IF bReset
     AND bError
THEN
	udnErrorNo := 0;					(* Error number *)
	sErrorMsg := ''; 					(* Error message *)
	tonWatchDog(IN := FALSE);

END_IF

(* Check inputs  *)
rtHandOn(CLK := bHandOn);
rtAutoOn(CLK := bAutoOn AND bReleaseOn AND bReleasePowerOn);
rtAutoOff(CLK := bAutoOff);

(* Check operating mode *)
IF bAutoHand					(* Automatic *)
THEN
	IF rtAutoOff.Q
	THEN
		bPowerOn := FALSE;

	ELSIF rtAutoOn.Q
		    AND bReleasePowerOn
	THEN
		bPowerOn := TRUE;
	END_IF;

ELSE						(* Manual *)
	IF rtHandOn.Q
	THEN
		IF bPowerOn
		THEN
			bPowerOn := FALSE;

		ELSIF bReleaseOn
			   AND bReleasePowerOn
		THEN
			bPowerOn := TRUE;
		END_IF
	END_IF

END_IF;

(* Timer starts when cylinder is not  in base and work position *)
tonWatchDog(
	IN := bPowerOn
		 AND bPowerSupplyOn
		 AND NOT bReady,
	PT := tTimeOut + tReadyDelay
);

(* Error if cylinder does not reach base or work position*)
IF tonWatchDog.Q
   AND NOT bError
THEN
	IF bPowerOn AND NOT bReady
	THEN
		udnErrorNo := 1; 								(* Set error number *)
		sErrorMsg := 'Not ready error';
	END_IF
END_IF

tonPowerSupplyOn(
	IN := bNoEStop
		 AND NOT bPowerSupplyOn,
	PT := tTimeOut
);

IF tonPowerSupplyOn.Q
THEN
	udnErrorNo := 2; 								(* Set error number *)
	sErrorMsg := 'Power supply error';
END_IF
(*
IF lrSetTemp > 0
     AND lrActTemp > lrMaxTemp
THEN
	udnErrorNo := 2; 								(* Set error number *)
	sErrorMsg := 'Temperatur over range';
END_IF
*)

bError := udnErrorNo <> 0;

fbReadyDelay(
	bEnable := TRUE,
	bIn := bPowerOn,
	tDelay := tReadyDelay
);

IF lrSetTemp <> 0
     AND bAutoHand 			(* Automatic *)
THEN
	bReady := bPowerOn
			   AND lrActTemp >= lrSetTemp;
ELSE
	bReady := fbReadyDelay.bOut;
END_IF

(* Scaling power *)
fbScalingSP(
	bEnable := TRUE,
	lrInput := lrSPPower, (* [%] *)
	lrXLowLimit := 0, (* [%] *)
	lrXUpperLimit := 100, (* [%] *)
	lrYLowLimit := lrPowerMin, (* 16#0000 = 0 [V] *)
	lrYUpperLimit := lrPowerMax, (* 16#7FFF = 10 [V] *)
	usiPrecision := 2
);
unCVPower := LREAL_TO_UINT(fbScalingSP.lrOutputPV);

END_FUNCTION_BLOCK

// ---- POUs/Tc2 Objects/Automation/NCiChannel/FB_CfgAxisInExt3DGroup.TcPOU
FUNCTION_BLOCK FB_CfgAxisInExt3DGroup
(*

The function block used to detects if are axis in a group or if the group is occupied. 

Constructor: 		Patryk Panylo
Company:		E. Riexinger GmbH
Date:			23.04.2015
Version:			1.00

Date:			Revision:		Who:				Comment
dd.mm.yyyy		x.xx			Initials			comment

*)
VAR_INPUT
	(* Input variables / Eingang Variablen *)
	bEnable						:BOOL;			(* Signal FB enable *)
	bExecute					:BOOL; 			(* Execute the programm *)
	udnGrpId						:UDINT;			(* Id of the 3D Group *)
	tTimeOut						:TIME := T#5s;	(* TimeOut *)
END_VAR
VAR_OUTPUT
	(* Output variables / Ausgang Variablen *)
	bGrpOccupied				:BOOL;			(* Axis in group detected *)
	bGrpEmpty					:BOOL;			(* Axis not in group detected *)
	bDone						:BOOL;			(* Command done *)
	bBusy						:BOOL;			(* Command busy *)
	bError						:BOOL;			(* Command error  *)
	udnErrorNo					:UDINT;			(* Error number *)
	sErrorMsg					:STRING; 		(* Error message *)
END_VAR
VAR_IN_OUT
	(* Input Output variables / Ausgang Variablen *)

END_VAR
VAR
	(* Enummerations *)
	etCfgAxisInExt3DGrp			:ET_CfgAxisInExt3DGroup;

	(* Variables *)
	stExt3dGrp 					:NCI_EXT3DGROUP;				(* Contains the Axis ID's *)

	bFirstTime					:BOOL;

	(* References *)

	(* Interfaces *)

	(* Instances *)
	fbCfgReadExt3DAxisIds		:CfgReadExt3DAxisIds;				(* The block CfgReadExt3DAxisIds reads the axis configuration of the advanced 3D group. *)

END_VAR

IF NOT bEnable
THEN
	bGrpOccupied := FALSE;			(* Axis in group detected *)
	bGrpEmpty :=FALSE;				(* Axis not in group detected *)
	bDone := FALSE;					(* Program done *)
	bBusy := FALSE;                                  	(* Program not busy *)
	bError := FALSE;                                 	(* Program not error *)
	udnErrorNo := 0;					(* Error number *)
	sErrorMsg := ''; 					(* Error message *)

	bFirstTime := FALSE;
	RETURN;
END_IF;

IF NOT bFirstTime
THEN
	bGrpOccupied := FALSE;			(* Axis in group detected *)
	bGrpEmpty :=FALSE;				(* Axis not in group detected *)
	bDone := FALSE;                                 	(* Program done *)
	bBusy := FALSE;                                  	(* Program not busy *)
	bError := FALSE;                                 	(* Program not error *)
	udnErrorNo := 0;					(* Error number *)
	sErrorMsg := ''; 					(* Error message *)

	fbCfgReadExt3DAxisIds(
		bExecute := FALSE,
		stExt3dGroup := stExt3dGrp
	);

	etCfgAxisInExt3DGrp := ET_CfgAxisInExt3DGrp_eWaitExecute;       				(* Next step *)
	
	bFirstTime := TRUE;
END_IF;

CASE etCfgAxisInExt3DGrp OF
        
	ET_CfgAxisInExt3DGrp_eWaitExecute:
		bBusy := FALSE;                                     		(* Program not busy *)
		bError := FALSE;                                    		(* Program not error *)

		IF bExecute
		THEN
			bDone := FALSE;                                 	(* Program done, in position *)
			bBusy := TRUE;                                  	(* Program busy *)
			udnErrorNo := 0;					(* Error number *)
			sErrorMsg := ''; 					(* Error message *)
	           
			etCfgAxisInExt3DGrp := ET_CfgAxisInExt3DGrp_eReadExt3DAxisIds;         		(* Next step *)
		END_IF;

	ET_CfgAxisInExt3DGrp_eReadExt3DAxisIds:

		fbCfgReadExt3DAxisIds(			(* Read axis ID's *)
			bExecute := TRUE ,
			nGroupId := udnGrpId,
			tTimeOut := tTimeOut,
			stExt3dGroup := stExt3dGrp
		);

		IF NOT fbCfgReadExt3DAxisIds.bBusy
		     AND NOT fbCfgReadExt3DAxisIds.bErr
		THEN
			fbCfgReadExt3DAxisIds(
				bExecute := FALSE,
				stExt3dGroup := stExt3dGrp
			);

			bGrpEmpty :=	stExt3dGrp.nXAxisId = 0						(* Check if axis in Group *)
						AND stExt3dGrp.nYAxisId = 0
						AND stExt3dGrp.nZAxisId = 0
						AND stExt3dGrp.nQ1AxisId =  0
						AND stExt3dGrp.nQ2AxisId =  0
						AND stExt3dGrp.nQ3AxisId =  0
						AND stExt3dGrp.nQ4AxisId =  0
						AND stExt3dGrp.nQ5AxisId =  0;
			bGrpOccupied := NOT bGrpEmpty ;
			
			etCfgAxisInExt3DGrp := ET_CfgAxisInExt3DGrp_eDone;            			(* Next step *)

		ELSIF fbCfgReadExt3DAxisIds.bErr
		THEN
			udnErrorNo := fbCfgReadExt3DAxisIds.nErrId;						(* Set error number *)

			fbCfgReadExt3DAxisIds(
				bExecute := FALSE,
				stExt3dGroup := stExt3dGrp
			);

			etCfgAxisInExt3DGrp := ET_CfgAxisInExt3DGrp_eError;            			(* Next step *)
		
		END_IF

	ET_CfgAxisInExt3DGrp_eDone:
		bDone := TRUE;                                      		(* Program done, in position *)
		bBusy := FALSE;                                     		(* Program not busy *)
	
		etCfgAxisInExt3DGrp := ET_CfgAxisInExt3DGrp_eNoExecute;            		(* Next step *)
	
	ET_CfgAxisInExt3DGrp_eError:
		bDone := FALSE;                                    	 	(* Program done, in position *)
		bError := TRUE;                                     		(* Program error *)
		bBusy := FALSE;                                     		(* Program not busy *)

		etCfgAxisInExt3DGrp := ET_CfgAxisInExt3DGrp_eNoExecute;            		(* Next step *)
	
	ET_CfgAxisInExt3DGrp_eNoExecute:
		IF NOT bExecute
		THEN
			bDone := FALSE;                                 	(* Program done *)
			bBusy := FALSE;                                 	(* Program not busy *)
			bError := FALSE;                                		(* Program not error *)

			etCfgAxisInExt3DGrp := ET_CfgAxisInExt3DGrp_eWaitExecute;       		(* Next step *)
	
		END_IF;
        
END_CASE;

END_FUNCTION_BLOCK

// ---- POUs/Tc2 Objects/Automation/Sawband/FB_Sawband.TcPOU
FUNCTION_BLOCK FB_Sawband
(*

The function block used to control the saw.

Constructor: 		Patryk Panylo
Company:		E. Riexinger GmbH
Date:			04.11.2015
Version:			1.00

Date:			Revision:		Who:				Comment
dd.mm.yyyy		x.xx			Initials			comment

*)
VAR_INPUT
	(* Input variables / Eingang Variablen *)
	bEnable					:BOOL;						(* Enable FB signal *)
	bNoEStop				:BOOL;						(* No ermergency Stop / Keine Notaus *)
	bAirPressure				:BOOL;						(* Signal air pressure *)
	bAutoHand				:BOOL;						(* Auto := TRUE, Hand := FALSE *)
	bHandStart				:BOOL;						(* Sawband hand start *)
	bHandStop				:BOOL;						(* Sawband hand stop *)
	bAutoStart				:BOOL;						(* Sawband auto start *)
	bAutoStop				:BOOL;						(* Sawband auto stop *)
	bSawbandAir				:BOOL;						(* Sawband air on *)
	bSawbandCtrlOK			:BOOL;						(* Sawband controller ok *)
	bSawbandNOK			:BOOL;						(* Sawband error *)
	udnIncEnc				:UDINT;						(* Value of encoder increment *)
	udnScalingDenom			:UDINT := 1;	  				(* Denominator for the conversion factor at the conversion of bus data to technical units [INC] *)
	lrScalingNum				:LREAL := 1.0;  				(* Numerator for the conversion factor at the conversion of bus data to technical units [technical units] *)
	lrTaskCycle				:LREAL := 0.002;				(* Cycle time of the task [sec], 0.002[s] => 2ms *)
	lrSawbandRefVelo		:LREAL := 1.0;					(* Referenc velocity of sawband [technical units/s]*)
	tSawbandCtrlOnDelay		:TIME := t#3s;					(* Sawband on delay *)
	tSawbandAirOffDelay		:TIME := t#10s;				(* Sawband air off delay *)
	tSawbandReadyDelay		:TIME := t#5s;					(* Sawband ready delay *)
END_VAR
VAR_OUTPUT
	(* Output variables / Ausgang Variablen *)
	bSawbandReady			:BOOL;						(* Sawband ready *)
	bSawbandCtrlOn			:BOOL;						(* Sawband controller on *)
	bSawbandAirOn			:BOOL;						(* Sawband air on*)
	bNotMoving				:BOOL;						(* Axis not moving *)
	lrActPosition				:LREAL;						(* Actual position [mm] *)
	lrActVelocity				:LREAL;						(* Actual velocity [mm/s] *)
	bError					:BOOL;						(* Error *)
	udnErrorNo				:UDINT;
	udnMessageNo			:UDINT;
	sMsg					:STRING;
END_VAR
VAR_IN_OUT

END_VAR
VAR
	(* Enummerations *)

	(* Variables *)
	stEncoderConfig				:ST_EncoderConfig;			(* Encoder configuration *)
	stAxis						:ST_AXIS_REF_V2;			(* The AXIS_REF data type  is an interface between the PLC and the NC and contains axis information *)
	bFirstTime					:BOOL;						(* First cycle *)

	(* References *)

	(* Interfaces *)

	(* Instances *)
	rtHandStart				:R_TRIG;
	rtHandStop				:R_TRIG;
	rtAutoStart				:R_TRIG;
	rtAutoStop				:R_TRIG;
	tonSawbandCtrlOnDelay	:TON;						(* Timer to delay *)
	tofSawbandAirOffDelay		:TOF;						(* Timer to delay *)
	tonSawbandReadyDelay  	:TON;						(* Timer to delay *)

	fbPositionEncoder			:FB_PositionEncoder;
END_VAR

IF NOT bEnable
THEN
	bSawbandCtrlOn := FALSE;
	bSawbandAirOn := FALSE;
	bError := FALSE;
	udnErrorNo := 0;
	udnMessageNo := 0;
	sMsg := '';
	tonSawbandCtrlOnDelay(IN := FALSE,
					       	    PT := tSawbandCtrlOnDelay);
	tofSawbandAirOffDelay(IN := FALSE,
	            			 	 PT := tSawbandAirOffDelay);
	tonSawbandReadyDelay(IN := FALSE,
					       		PT := tSawbandReadyDelay);
	bFirstTime := FALSE;
    RETURN;
END_IF;

IF NOT bFirstTime
THEN
	bError := FALSE;
	udnErrorNo := 0;
	udnMessageNo := 0;
	sMsg := '';
	tonSawbandCtrlOnDelay(IN := FALSE,
					       	    PT := tSawbandCtrlOnDelay);
	tofSawbandAirOffDelay(IN := FALSE,
	            			 	 PT := tSawbandAirOffDelay);
	tonSawbandReadyDelay(IN := FALSE,
					       		PT := tSawbandReadyDelay);
	bFirstTime := TRUE;
END_IF;

(* Start / Stop sawband *)
rtHandStart(CLK := bHandStart);
rtHandStop(CLK := bHandStop);
rtAutoStart(CLK := bAutoStart);
rtAutoStop(CLK := bAutoStop);

IF rtHandStop.Q
     OR rtAutoStop.Q
     OR NOT bNoEStop
     OR bSawbandNOK
THEN
	tofSawbandAirOffDelay.IN := FALSE;;
	tonSawbandCtrlOnDelay.IN := FALSE;

ELSIF SEL(bAutoHand, rtHandStart.Q, rtAutoStart.Q)
	    AND bNoEStop
	    AND bAirPressure
	    AND NOT bSawbandNOK
THEN
	tofSawbandAirOffDelay.IN := TRUE;;
	tonSawbandCtrlOnDelay.IN := TRUE;

END_IF

(* Sawband air stop after delay *)
tofSawbandAirOffDelay(
         PT := tSawbandAirOffDelay
);

bSawbandAirOn := tofSawbandAirOffDelay.Q
				OR ( NOT bAutoHand
					AND bSawbandAir);

(* Sawband controller on after delay *)
tonSawbandCtrlOnDelay(
         PT := tSawbandCtrlOnDelay
);

bSawbandCtrlOn := tonSawbandCtrlOnDelay.Q;

(* Sawband ready after delay *)
tonSawbandReadyDelay(
	IN := bSawbandCtrlOn,
	PT := tSawbandReadyDelay
);

A_PositionDynamics();
A_Alarm();

bSawbandReady := bSawbandCtrlOK
				   AND NOT bSawbandNOK
				   AND NOT bNotMoving
				   AND NOT bError
				   AND lrActVelocity >= lrSawbandRefVelo
				   AND tonSawbandReadyDelay.Q;

ACTION A_Alarm:

(* Check error *)
IF bSawbandNOK
THEN
	udnErrorNo := 1;
	udnMessageNo := 0;
	sMsg := 'Sawband nok signal';

ELSIF (NOT bSawbandCtrlOK
	    	      OR bNotMoving)
	   AND tonSawbandReadyDelay.Q
THEN
	udnErrorNo := 2;
	udnMessageNo := 0;
	sMsg := 'Sawband not ready';

ELSE
	udnErrorNo := 0;
	udnMessageNo := 0;
	sMsg := '';

END_IF

bError := udnErrorNo > 0;
END_ACTION

ACTION A_PositionDynamics:

(* Position encoding *)
stEncoderConfig.etScalingMethod := ET_ScalingMethod_eSMLinear;
stAxis.stScaling.etScalingMethod := ET_ScalingMethod_eSMLinear;
stAxis.stScaling.lrTaskCycle := lrTaskCycle;
stAxis.stScaling.udnScalingDenom := udnScalingDenom; (* inc *)
stAxis.stScaling.lrScalingNum := lrScalingNum; (* mm *)

fbPositionEncoder(
	bEnable := TRUE,
	dwEncCurrentValue := udnIncEnc,
	stEncCfg := stEncoderConfig,
	pAxis := ADR(stAxis)
);

lrActPosition := fbPositionEncoder.pAxis^.stPosition.lrActPos / 1000 (* m *);
lrActVelocity := fbPositionEncoder.pAxis^.stDynamics.lrActVelo * 60 (* mm/min *);

bNotMoving := FALSE;

IF lrActVelocity = 0.0
THEN
	bNotMoving := TRUE;
END_IF
END_ACTION

END_FUNCTION_BLOCK

// ---- POUs/Tc2 Objects/Automation/Spindle/FB_CoolingDevice.TcPOU
FUNCTION_BLOCK FB_CoolingDevice
(*

The function block used to control power supply.

Constructor: 		Patryk Panylo
Company:		E. Riexinger GmbH
Date:			23.04.2015
Version:			1.00

Date:			Revision:		Who:				Comment
dd.mm.yyyy		x.xx			Initials			comment

*)
VAR_INPUT
	(* Input variables / Eingang Variablen *)
	bEnable					:BOOL;						(* Enable FB signal *)
	bIn						:BOOL;						(* Input signal *)
	tCoolingDeviceOn			:TIME := t#2s;					(* Timeout power supply on *)
	tCoolingDeviceOff			:TIME := t#1s;					(* Timeout power supply off *)
END_VAR
VAR_OUTPUT
	(* Output variables / Ausgang Variablen *)
	bOut					:BOOL;						(* Air pressure ok *)
	bError					:BOOL;						(* Error by no air pressure *)
	udnErrorNo				:UDINT;
	udnMessageNo			:UDINT;
	sMsg					:STRING;
END_VAR
VAR_IN_OUT

END_VAR
VAR
	(* Enummerations *)

	(* Variables *)
	bFirstTime				:BOOL;						(* First cycle *)

	(* References *)

	(* Interfaces *)

	(* Instances *)
	tonCoolingDeviceOn		:TON;						(* Timer to delay *)
	tofCoolingDeviceOff		:TOF;						(* Timer to delay *)
	tCoolingDevice			:BOOL;
END_VAR

IF NOT bEnable
THEN
	bOut := TRUE;
	bError := FALSE;
	udnErrorNo := 0;
	udnMessageNo := 0;
	sMsg := '';
	tonCoolingDeviceOn(IN := FALSE,
				            PT := tCoolingDeviceOn);
	tofCoolingDeviceOff(IN := FALSE,
	            			 PT := tCoolingDeviceOff);
	bFirstTime := FALSE;
    RETURN;
END_IF;

IF NOT bFirstTime
THEN
	bError := FALSE;
	udnErrorNo := 0;
	udnMessageNo := 0;
	sMsg := '';
	tonCoolingDeviceOn(IN := FALSE,
	          			  PT := tCoolingDeviceOn);
	tofCoolingDeviceOff(IN := FALSE,
	             			 PT := tCoolingDeviceOff);
	bFirstTime := TRUE;
END_IF;

(* Timer starts when came rising edge of signal *)
tonCoolingDeviceOn(
	IN := bIn,
         PT := tCoolingDeviceOn
);

tofCoolingDeviceOff(
	IN := bIn,
         PT := tCoolingDeviceOff
);

bOut := tonCoolingDeviceOn.Q;
bError := NOT tofCoolingDeviceOff.Q;

IF bError
THEN
	udnErrorNo := 1;
	udnMessageNo := 0;
	sMsg := 'No power supply';
ELSE
	udnErrorNo := 0;
	udnMessageNo := 0;
	sMsg := '';
END_IF;

END_FUNCTION_BLOCK

// ---- POUs/Tc2 Objects/Automation/Spindle/FB_SpindlePreheat.TcPOU
FUNCTION_BLOCK FB_SpindlePreheat
(*

The function block used to start spindle preheat procedure.

Constructor: 		Patryk Panylo
Company:		E. Riexinger GmbH
Date:			26.06.2015
Version:			1.00

Date:			Revision:		Who:				Comment
dd.mm.yyyy		x.xx			Initials			comment

*)
VAR_INPUT
	(* Input variables / Eingang Variablen *)
	bEnable						:BOOL;						(* Enable FB signal *)
	bNoEmergencyStop			:BOOL;						(* NotAus signal *)
	bExecute					:BOOL;						(* Spindle start *)
	bInterrupt						:BOOL;						(* Interrupt *)
	bPlusRelease				:BOOL;						(* Plus move release *)
	bMinusRelease				:BOOL;						(* Minus move release *)
	bReset						:BOOL;						(* Reset procedure*)
	bCtrlEnabled					:BOOL;						(* Controller enabled *)
	bSetNewSpdlPreheat			:BOOL;						(* Set new spindle preheat *)
	bSetDailyPreheat				:BOOL;						(* Set daily preheat *)
	tSetPeriod					:TIME;						(* Set period time *)
	lrMaxRpm					:LREAL;						(* Max rpm [U/min]  *)
	bRpmIsZero					:BOOL;						(* Spindle standstill *)
	bRpmReached				:BOOL;						(* Spindle speed reached *)
END_VAR
VAR_OUTPUT
	(* Output variables / Ausgang Variablen *)
	bValid						:BOOL;						(* Preheat valid *)
	unSpindleDurationPercent		:UINT;						(* Actual spindle duration in percent*)
	bControlerOn					:BOOL;						(* Controler on *)
	bDone						:BOOL;						(* Program done *)
	bBusy						:BOOL;						(* Program busy *)
	bError						:BOOL;						(* Program error *)
	udnErrorNo					:UDINT;						(* Error number *)
	sErrorMsg					:STRING;
END_VAR
VAR_IN_OUT
	(* Input Output variables / Ausgang Variablen *)
	Axis							:AXIS_REF;					(* The AXIS_REF data type  is an interface between the PLC and the NC and contains axis information *)
	arstPhasesNewSpdl			:ARRAY [1..ungGr05MaxPhasesNewSpdl] OF ST_SpindlePreheat; 				(* Starting new spindel phases *)
	arstPhasesDailyPreheat		:ARRAY [1..ungGr05MaxPhasesDailyPreheat] OF ST_SpindlePreheat; 			(* Starting daily preheat phases *)
END_VAR
VAR
	(* Enummerations *)
	etSpindlePreheat				:ET_SpindlePreheat;				(* Spindle  mode enum variable *)

	(* Variables *)
	otstTime						:OTSTRUCT;						(* Time in OTSTRUCT *)
	unPhase						:UINT;							(* Phase counter *)
	lrSpdlTimeAsHour				:LREAL;							(* The running time of spindle procedures [h] *)
	lrStartSpdlProcTimeAsHour		:LREAL;							(* Start time of spindle procedure [h] *)
	lrSystemNewTimeAsHour 		:LREAL; 							(* System Time [h] *)
	lrPeriodAsHour				:LREAL; 							(* Period Time [h] *)
	lrWeekAsHour				:LREAL;							(* Week [h] *)
	lrDayAsHour					:LREAL;							(* Day [h] *)
	lrHour						:LREAL;							(* Hour [h] *)
	lrMinuteAsHour				:LREAL;							(* Minute Time [h] *)
	lrSecondAsHour				:LREAL;							(* Second Time [h] *)
	lrMillisecondAsHour			:LREAL;							(* Millisecond Time [h] *)

	bNewSpdl					:BOOL; 							(* New spindel phases *)
	bDailyPreheat				:BOOL; 							(* Daily preheat phases *)

	bFirstTime					:BOOL;

	(* References *)

	(* Interfaces *)

	(* Instances *)
	fbGetSystemTime				:GETSYSTEMTIME;				(* Detects System time *)
	rtReset						:R_TRIG; 						(* Positive edge for reset procedure *)
	rtExecute						:R_TRIG;							(* Positive edge for execute *)
	tonDuration					:TON;
	fbMCMoveVelo				:MC_MoveVelocity;
	fbMCStop					:MC_Stop;
	tonCtrlEnabled				:TON;
	rtSetNewSpdlPreheat			:R_TRIG;							(* Set new spindle preheat *)
	rtSetDailyPreheat				:R_TRIG;							(* Set daily preheat *)
END_VAR
VAR PERSISTENT
	lrSystemOldTimeAsHour 		:LREAL; 						(* System Time [h] *)
	bProcInterrupted				:BOOL;						(* Statring procedure interupted *)
END_VAR


IF NOT bEnable						(* Signal FB enable *)
THEN
	bValid := FALSE;;					(* Preheat valid *)
	bControlerOn := FALSE;			(* Controler off *)
	bDone := FALSE;					(* Program done *)
	bBusy := FALSE;                                  	(* Program not busy *)
	bError := FALSE;                                 	(* Program not error *)
	udnErrorNo := 0;                                 		(* Error number *)

	tonCtrlEnabled(IN := FALSE);

	bFirstTime := FALSE;

	RETURN;
END_IF;

(* Calculate system time *)
fbGetSystemTime();
lrSystemNewTimeAsHour := UINT64_TO_LREAL(IN := ULARGE_INTEGER(
	dwHighPart := fbGetSystemTime.timeHiDW,
	dwLowPart := fbGetSystemTime.timeLoDW))
	/ 10				(* Calculate into mycro seconds *)
	/ 1000			(* Calculate into millis econds *)
	/ 1000			(* Calculate into seconds *)
	/ 60				(* Calculate into minutes *)
	/ 60;				(* Calculate into hours *)

(* Calculate period time *)
otstTime := TIME_TO_OTSTRUCT(TIN := tSetPeriod);

lrWeekAsHour := otstTime.wWeek * 168.0;						(* Calculate into hours*)
lrDayAsHour := otstTime.wDay * 24.0;							(* Calculate into hours *)
lrHour := otstTime.wHour ;
lrMinuteAsHour := otstTime.wMinute  / 60.0;						(* Calculate into hours *)
lrSecondAsHour := otstTime.wSecond / 3600.0;					(* Calculate into hours *)
lrMillisecondAsHour := otstTime.wMilliseconds / 3600000.0 ;		(* Calculate into hours *)

lrPeriodAsHour :=  lrWeekAsHour							(* Calculate period *)
				+ lrDayAsHour
				+ lrHour
				+ lrMinuteAsHour
		 		+ lrSecondAsHour
				+ lrMillisecondAsHour;

(* Save last time activated of spindle *)
IF NOT Axis.NcToPlc.StateDWord.2			(* Axis moving *)
    AND Axis.NcToPlc.SetVelo <> 0.0
    AND NOT bProcInterrupted
    AND NOT bBusy
THEN
	lrSystemOldTimeAsHour := lrSystemNewTimeAsHour;
END_IF

rtSetNewSpdlPreheat(CLK := bSetNewSpdlPreheat);
rtSetDailyPreheat(CLK := bSetDailyPreheat);

IF rtSetNewSpdlPreheat.Q
THEN
	lrSystemOldTimeAsHour := 0.0;
ELSIF rtSetDailyPreheat.Q
	    AND lrSystemOldTimeAsHour <> 0
THEN
	lrSystemOldTimeAsHour := 1.0;
END_IF

rtReset (CLK := bReset);											(* Positive edge for reset procedure*)
IF rtReset.Q
     AND bError
THEN
	bControlerOn := FALSE;				(* Controler off *)
	bDone := FALSE;					(* Program done *)
	bBusy := FALSE;                                  	(* Program not busy *)
	bError := FALSE;                                 	(* Program not error *)
	udnErrorNo := 0;                                 		(* Error number *)

	(* The function block MC_MoveVelocity starts a continuous movement with specified velocity and direction.  *)
	fbMCMoveVelo(
		Execute := FALSE,
		Axis := Axis,
	 );

	(* The function block MC_Stop stops an axis with a defined braking ramp and blocks the axis for any motion commands.  *)
	fbMCStop(
		Execute := FALSE,
		Axis := Axis,
	);

	tonDuration(IN:= FALSE);

	etSpindlePreheat := ET_SpindlePreheat_eWaitExecute;       			(* Next step *)

END_IF

(* Positive edge for execute *)
rtExecute(CLK := bExecute);
IF rtExecute.Q
THEN
	tonCtrlEnabled(IN := FALSE);

	bControlerOn := bMinusRelease
     				   AND bPlusRelease
     				   AND bNoEmergencyStop
     				   AND NOT bInterrupt;

	IF lrSystemNewTimeAsHour - lrSystemOldTimeAsHour < lrPeriodAsHour
	THEN
		bControlerOn := FALSE;
		bValid := TRUE;
	ELSE
		bValid := FALSE;
	END_IF

	RETURN;
ELSE
	tonCtrlEnabled(IN := bControlerOn
					   AND NOT bCtrlEnabled,
				   PT := t#3s);

	IF NOT bControlerOn
	     OR NOT bCtrlEnabled
	THEN
		bBusy := FALSE;                                 	(* Program not busy *)

		IF tonCtrlEnabled.Q
		THEN
			bControlerOn := FALSE;
		END_IF

		RETURN;
	ELSE
		tonCtrlEnabled(IN := FALSE);
	END_IF
END_IF;

IF NOT bCtrlEnabled
     OR NOT bNoEmergencyStop
     OR NOT bMinusRelease
     OR NOT bPlusRelease
     OR bInterrupt
THEN
	bControlerOn := FALSE;			(* Controler off *)

	(* Interrupt only when procedure has been busy  *)
	IF bBusy
	     AND NOT bProcInterrupted
	THEN
		bBusy := FALSE;                                 	(* Program not busy *)
		bProcInterrupted := TRUE;
	END_IF

	IF Axis.NcToPlc.StateDWord.2			(* Axis not moving *)
	THEN
		unSpindleDurationPercent := 0;
	END_IF

	bFirstTime := FALSE;

	RETURN;
END_IF

IF NOT bFirstTime
THEN
	bDone := FALSE;                                	(* Program done *)
	bBusy := FALSE;                                 	(* Program not busy *)
	bError := FALSE;                                 	(* Program not error *)
	udnErrorNo := 0;                                 		(* Error number *)

	(* The function block MC_MoveVelocity starts a continuous movement with specified velocity and direction.  *)
	fbMCMoveVelo(
		Execute := FALSE,
		Axis := Axis,
	 );

	(* The function block MC_Stop stops an axis with a defined braking ramp and blocks the axis for any motion commands.  *)
	fbMCStop(
		Execute := FALSE,
		Axis := Axis,
	);

	tonDuration(IN:= FALSE);

	etSpindlePreheat := ET_SpindlePreheat_eWaitExecute;       			(* Next step *)

	bFirstTime := TRUE;
END_IF;

IF bBusy
     AND Axis.NcToPlc.SetVelo <> 0.0
     AND NOT Axis.NcToPlc.StateDWord.2			(* Axis moving *)
THEN
	IF lrSystemNewTimeAsHour - lrStartSpdlProcTimeAsHour >= lrSpdlTimeAsHour
	THEN
		lrStartSpdlProcTimeAsHour := lrSystemNewTimeAsHour;
		IF unSpindleDurationPercent < 100
		THEN
			unSpindleDurationPercent := unSpindleDurationPercent + 1;
		ELSE
			unSpindleDurationPercent := 100;
		END_IF
	END_IF
ELSE
	IF Axis.NcToPlc.StateDWord.2			(* Axis not moving *)
	THEN
		unSpindleDurationPercent := 0;
	END_IF
END_IF

CASE etSpindlePreheat OF

	ET_SpindlePreheat_eWaitExecute:
		bBusy := FALSE;                                     		(* Program not busy *)
		bError := FALSE;                                    		(* Program not error *)

		bNewSpdl := FALSE; 					(* New spindel phases *)
		bDailyPreheat := FALSE; 				(* Daily preheat phases *)

		IF bControlerOn
		    AND bCtrlEnabled
		THEN
			bDone := FALSE;						(* Command done *)
			bBusy := TRUE;						(* Command busy *)
			bError := FALSE;						(* Command error  *)
			udnErrorNo := 0;						(* Error number *)
			sErrorMsg := ''; 						(* Error message *)

			tonDuration(IN:= FALSE);
			lrSpdlTimeAsHour := 0.0;

			(* New spindle starting procedure *)
			IF lrSystemOldTimeAsHour = 0
			THEN

				FOR unPhase := 1 TO ungGr05MaxPhasesNewSpdl
				DO
					(* Convert  duration time to OTSTRUCT*)
					arstPhasesNewSpdl[unPhase].otstDuration := TIME_TO_OTSTRUCT(TIN := arstPhasesNewSpdl[unPhase].tDuration);

					(* Calculate period time *)
					lrWeekAsHour := arstPhasesNewSpdl[unPhase].otstDuration.wWeek * 168.0;						(* Calculate into hours*)
					lrDayAsHour := arstPhasesNewSpdl[unPhase].otstDuration.wDay * 24.0;							(* Calculate into hours *)
					lrHour := arstPhasesNewSpdl[unPhase].otstDuration.wHour;
					lrMinuteAsHour := arstPhasesNewSpdl[unPhase].otstDuration.wMinute  / 60.0;						(* Calculate into hours *)
					lrSecondAsHour := arstPhasesNewSpdl[unPhase].otstDuration.wSecond / 3600.0;					(* Calculate into hours *)
					lrMillisecondAsHour := arstPhasesNewSpdl[unPhase].otstDuration.wMilliseconds / 3600000.0 ;			(* Calculate into hours *)

					lrSpdlTimeAsHour :=  lrSpdlTimeAsHour														(* Calculate period *)
									      + lrWeekAsHour
									      + lrDayAsHour
							 	    	      + lrHour
									      + lrMinuteAsHour
							 	    	      + lrSecondAsHour
									      + lrMillisecondAsHour;

					(* Set Limited Override *)
					arstPhasesNewSpdl[unPhase].dwOverride := LIMIT(
						0,														(* Min 0 [%]  override*)
						arstPhasesNewSpdl[unPhase].dwOverride,					(* Current [%] override*)
						100														(* Max 100 [%] override *)
					);

					(* Set Speed *)
					arstPhasesNewSpdl[unPhase].dwSpeedRpm := (LREAL_TO_DWORD(lrMaxRpm) * arstPhasesNewSpdl[unPhase].dwOverride)/100;				(* Current RPM [U/min] *)

				END_FOR

				lrSpdlTimeAsHour := lrSpdlTimeAsHour / 100.0; 				(* Normalized to [%]*)
				lrStartSpdlProcTimeAsHour := lrSystemNewTimeAsHour;

				unPhase := 1;
				bBusy := TRUE;				(* Program Busy *)
				bNewSpdl := TRUE; 					(* New spindel phases *)
				bProcInterrupted := FALSE;

				etSpindlePreheat := ET_SpindlePreheat_eStartNewSpindle;		(* Next step *)

			(* Daily preheat starting procedure *)
			ELSIF lrSystemNewTimeAsHour - lrSystemOldTimeAsHour > lrPeriodAsHour
			THEN

				FOR unPhase := 1 TO ungGr05MaxPhasesDailyPreheat
				DO
					(* Convert  duration time to OTSTRUCT*)
					arstPhasesDailyPreheat[unPhase].otstDuration := TIME_TO_OTSTRUCT(TIN := arstPhasesDailyPreheat[unPhase].tDuration);

					(* Calculate period time *)
					lrWeekAsHour := arstPhasesDailyPreheat[unPhase].otstDuration.wWeek * 168.0;						(* Calculate into hours*)
					lrDayAsHour := arstPhasesDailyPreheat[unPhase].otstDuration.wDay * 24.0;							(* Calculate into hours *)
					lrHour := arstPhasesDailyPreheat[unPhase].otstDuration.wHour ;
					lrMinuteAsHour := arstPhasesDailyPreheat[unPhase].otstDuration.wMinute  / 60.0;						(* Calculate into hours *)
					lrSecondAsHour := arstPhasesDailyPreheat[unPhase].otstDuration.wSecond / 3600.0;					(* Calculate into hours *)
					lrMillisecondAsHour := arstPhasesDailyPreheat[unPhase].otstDuration.wMilliseconds / 3600000.0 ;			(* Calculate into hours *)

					lrSpdlTimeAsHour :=  lrSpdlTimeAsHour															(* Calculate period *)
									     + lrWeekAsHour
									     + lrDayAsHour
							 	    	     + lrHour
									     + lrMinuteAsHour
							 	   	     + lrSecondAsHour
									     + lrMillisecondAsHour;

					(* Set Limited Override *)
					arstPhasesDailyPreheat[unPhase].dwOverride := LIMIT(
						0,														(* Min 0 [%]  override*)
						arstPhasesDailyPreheat[unPhase].dwOverride,				(* Current [%] override*)
						100														(* Max 100 [%] override *)
					);

					(* Set Speed *)
					arstPhasesDailyPreheat[unPhase].dwSpeedRpm := (LREAL_TO_DWORD(lrMaxRpm) * arstPhasesDailyPreheat[unPhase].dwOverride)/100;				(* Current RPM [U/min] *)

				END_FOR

				lrSpdlTimeAsHour := lrSpdlTimeAsHour / 100.0; 				(* Normalized to [%]*)
				lrStartSpdlProcTimeAsHour := lrSystemNewTimeAsHour;

				unPhase := 1;
				bBusy := TRUE;				(* Program Busy *)
				bDailyPreheat := TRUE; 				(* Daily preheat phases *)
				bProcInterrupted := FALSE;

				etSpindlePreheat := ET_SpindlePreheat_eStartDailyPreheat;		(* Next step *)

			END_IF;
		END_IF;

	ET_SpindlePreheat_eStartNewSpindle:
		fbMCMoveVelo.Velocity := arstPhasesNewSpdl[unPhase].dwSpeedRpm;				(* Set speed RPM [U/min] *)
		tonDuration.PT := arstPhasesNewSpdl[unPhase].tDuration;							(* Set duration time *)

		etSpindlePreheat := ET_SpindlePreheat_eStartSpindle;		(* Next step *)

	ET_SpindlePreheat_eStartDailyPreheat:
		fbMCMoveVelo.Velocity := arstPhasesDailyPreheat[unPhase].dwSpeedRpm;			(* Set speed RPM [U/min] *)
		tonDuration.PT := arstPhasesDailyPreheat[unPhase].tDuration;						(* Set duration time *)

		etSpindlePreheat := ET_SpindlePreheat_eStartSpindle;		(* Next step *)

	ET_SpindlePreheat_eStartSpindle:
		fbMCMoveVelo.Execute := TRUE;

		IF fbMCMoveVelo.Busy
		THEN
			etSpindlePreheat := ET_SpindlePreheat_eWfStartSpindle;         		(* Next step *)

		ELSIF fbMCMoveVelo.Error
		THEN
			fbMCMoveVelo.Execute := FALSE;

			etSpindlePreheat := ET_SpindlePreheat_eError;         		(* Next step *)

		END_IF

	ET_SpindlePreheat_eWfStartSpindle:
		IF fbMCMoveVelo.InVelocity
		     AND NOT fbMCMoveVelo.Error
		     AND Axis.NcToPlc.StateDWord.12					(* Constant velocity *)
		     AND bRpmReached
		THEN
			fbMCMoveVelo.Execute := FALSE;

			etSpindlePreheat := ET_SpindlePreheat_eWfStartSpindleProc;         		(* Next step *)

		ELSIF fbMCMoveVelo.Error
		THEN
			fbMCMoveVelo.Execute := FALSE;

			etSpindlePreheat := ET_SpindlePreheat_eError;         		(* Next step *)

		END_IF

	ET_SpindlePreheat_eWfStartSpindleProc:
		tonDuration(IN := TRUE);

		IF tonDuration.Q
		THEN
			tonDuration(IN:= FALSE);

			(* Phase incrementation *)
			unPhase := unPhase + 1;

			IF bNewSpdl
			    AND unPhase <= ungGr05MaxPhasesNewSpdl
			THEN
				fbMCMoveVelo.Velocity := arstPhasesNewSpdl[unPhase].dwSpeedRpm;				(* Set speed RPM [U/min] *)
				tonDuration.PT := arstPhasesNewSpdl[unPhase].tDuration;							(* Set duration time *)

				etSpindlePreheat := ET_SpindlePreheat_eStartSpindle;

			ELSIF bDailyPreheat
				   AND unPhase <= ungGr05MaxPhasesDailyPreheat
			THEN
				fbMCMoveVelo.Velocity := arstPhasesDailyPreheat[unPhase].dwSpeedRpm;			(* Set speed RPM [U/min] *)
				tonDuration.PT := arstPhasesDailyPreheat[unPhase].tDuration;						(* Set duration time *)

				etSpindlePreheat := ET_SpindlePreheat_eStartSpindle;

			ELSE
				etSpindlePreheat := ET_SpindlePreheat_eSpindleStop;

			END_IF
		END_IF

	ET_SpindlePreheat_eSpindleStop:
		fbMCStop.Execute := TRUE;
		fbMCMoveVelo.Velocity := 0.0;

		IF fbMCStop.Busy
		THEN
			etSpindlePreheat := ET_SpindlePreheat_eWfSpindleStopped;         		(* Next step *)

		ELSIF fbMCStop.Error
		THEN
			fbMCStop.Execute := FALSE;

			etSpindlePreheat := ET_SpindlePreheat_eError;         		(* Next step *)

		END_IF

	ET_SpindlePreheat_eWfSpindleStopped:
		IF fbMCStop.Done
		     AND NOT fbMCStop.Error
		     AND Axis.NcToPlc.StateDWord.2			(* Axis not moving *)
		     AND Axis.NcToPlc.SetVelo = 0.0
		     AND bRpmIsZero
		THEN
			fbMCStop.Execute := FALSE;

			etSpindlePreheat := ET_SpindlePreheat_eDone;         		(* Next step *)

		ELSIF fbMCStop.Error
		THEN
			fbMCStop.Execute := FALSE;

			etSpindlePreheat := ET_SpindlePreheat_eError;         		(* Next step *)

		END_IF

	ET_SpindlePreheat_eDone:
		bValid := TRUE;						(* Preheat valid *)
		bControlerOn := FALSE;				(* Controler off *)
		bDone := TRUE;                                     		(* Program done, in position *)
		bBusy := FALSE;                                     		(* Program not busy *)

		(* Save last time activated of the starting procedure *)
		lrSystemOldTimeAsHour := lrSystemNewTimeAsHour;

		etSpindlePreheat := ET_SpindlePreheat_eNoExecute;            	(* Next step *)

	ET_SpindlePreheat_eError:
		bDone := FALSE;                                     		(* Program done, in position *)
		bControlerOn := FALSE;				(* Controler off *)
		bError := TRUE;                                     		(* Program error *)
		bBusy := FALSE;                                     		(* Program not busy *)
	
		etSpindlePreheat := ET_SpindlePreheat_eNoExecute;           	(* Next step *)

	ET_SpindlePreheat_eNoExecute:
		IF NOT bExecute
		THEN
			bNewSpdl := FALSE; 				(* New spindel phases *)
			bDailyPreheat := FALSE; 			(* Daily preheat phases *)

			bControlerOn := FALSE;				(* Controler off *)
			bDone := FALSE;                                 	(* Program done *)
			bBusy := FALSE;                                		(* Program not busy *)
			bError := FALSE;                                		(* Program not error *)
		
			etSpindlePreheat := ET_SpindlePreheat_eWaitExecute;       (* Next step *)
		
		END_IF;

END_CASE;

(* The function block MC_MoveVelocity starts a continuous movement with specified velocity and direction.  *)
fbMCMoveVelo(
	Direction := MC_Positive_Direction, (* MC_Negative_Direction *)
	Axis := Axis
 );

(* The function block MC_Stop stops an axis with a defined braking ramp and blocks the axis for any motion commands.  *)
fbMCStop(
	Axis := Axis,
);

END_FUNCTION_BLOCK

// ---- POUs/Tc2 Objects/Automation/Spindle/FB_ToolStorage.TcPOU
FUNCTION_BLOCK FB_ToolStorage
(*

The function block used to storage the tool parameters.

Constructor: 		Patryk Panylo
Company:		E. Riexinger GmbH
Date:			18.06.2018
Version:			1.00

Date:			Revision:		Who:				Comment
dd.mm.yyyy		x.xx			Initials			comment

*)
VAR_INPUT
	(* Input variables / Eingang Variablen *)
	bEnable						:BOOL;						(* Enable FB signal *)
	bReset						:BOOL;						(* Reset *)
	bResetSelectedToolNest		:BOOL;						(* Reset selected tool nest *)
	unSelectedToolNest			:UINT;						(* Selected tool nest *)
	bResetAllToolNests			:BOOL;						(* Reset all tool nests  *)
	bExeToolNest				:BOOL;						(* Execute  tool nest *)
	unToolNo					:UINT;						(* Tool number *)
	bToolLifetimeOn				:BOOL;						(* Tool lifetime enabled *)
	rToolRotationalSpeedAct		:REAL;						(* Tool current rotational speed *)
	parbToolNestPresent			:POINTER TO ARRAY[0..unToolStorageCapacity] OF BOOL;				(* Tool in nest present *)
	parunToolNo					:POINTER TO ARRAY[0..unToolStorageCapacity] OF UINT;				(* Tool nummer *)
	parsToolDescription			:POINTER TO ARRAY[0..unToolStorageCapacity] OF STRING(11);		(* Tool description *)
	parunToolRotationalSpeed 		:POINTER TO ARRAY[0..unToolStorageCapacity] OF UINT;				(* Rotational speed *)
	parunToolLifetimeSet			:POINTER TO ARRAY[0..unToolStorageCapacity] OF UINT;				(* Setpoint tool lifetime *)
	parunToolLifetimeAct			:POINTER TO ARRAY[0..unToolStorageCapacity] OF UINT;				(* Curret tool lifetime *)
	paretToolStatus				:POINTER TO ARRAY[0..unToolStorageCapacity] OF ET_ToolStatus;		(* Tool status *)
	unToolNestUsingMax			:UINT;						(* Tool nest using maximal number *)
	tWatchdog					:TIME := t#5s;					(* Watchdog time *)
	lrTaskCycle					:LREAL;						(* Task cycle *)
END_VAR
VAR_OUTPUT
	(* Output variables / Ausgang Variablen *)
	bDone						:BOOL;						(* Program done *)
	bBusy						:BOOL;						(* Program busy *)
	bError						:BOOL;						(* Program error *)
	udnErrorNo					:UDINT;						(* Error number *)
END_VAR
VAR_IN_OUT
	unToolNestPrv				:UINT;												(* Previous tool nest number *)
	unToolNestAct				:UINT;												(* Current tool nest number *)
	unToolNestUsing				:UINT;												(* Using tool nest number *)
END_VAR
VAR
	(* Enummerations *)
	etToolStorage				:ET_ToolStorage;

	(* Variables *)
	unToolNestCount				:UINT;						(* Tool nest counter *)
	unToolNestSearchCount		:UINT;						(* Tool nest search counter  *)
	rToolLifetime					:REAL;						(* Tool lifetime *)
	bToolLifetimeReached			:BOOL;						(* Tool lifetime reached *)

	unIdxToolNestCount			:UINT;
	unLifetimeOnNewTool			:UINT;

	bFirstTime					:BOOL;						(* First cycle *)

	(* References *)

	(* Interfaces *)

	(* Instances *)
	rtResetSelectedToolNest		:R_TRIG;
	rtResetAllToolNests			:R_TRIG;
	rtExeToolNest				:R_TRIG;
	tonWatchdog					:TON;
END_VAR
VAR CONSTANT
	unToolStorageCapacity		:UINT := 32;
END_VAR

IF NOT bEnable
THEN
	bDone := FALSE;					(* Program done *)
	bBusy := FALSE;                                  	(* Program not busy *)
	bError := FALSE;                                 	(* Program not error *)
	udnErrorNo := 0;                                 		(* Error number *)

	tonWatchdog(IN := FALSE);

	etToolStorage := ET_ToolStorage_eWaitExecute;       				(* Next step *)

	bFirstTime := FALSE;
	RETURN;
END_IF;

IF NOT bFirstTime
THEN
	bDone := FALSE;					(* Program done *)
	bBusy := FALSE;                                  	(* Program not busy *)
	bError := FALSE;                                 	(* Program not error *)
	udnErrorNo := 0;                                 		(* Error number *)

	tonWatchdog(IN := FALSE);

	etToolStorage := ET_ToolStorage_eWaitExecute;       				(* Next step *)

	bFirstTime := TRUE;
END_IF;

IF unToolNestUsingMax > unToolStorageCapacity
THEN
	unToolNestUsingMax := unToolStorageCapacity;
END_IF

(* Get current tool *)
IF unToolNestCount >= unToolNestUsingMax
THEN
	unToolNestCount := 0;
END_IF
unToolNestCount := unToolNestCount + 1;

(* Control tool lifetime *)
IF parunToolLifetimeSet^[unToolNestCount] <> 0															(* If 0 then tool lifetime monitoring is not active *)
THEN
	IF parunToolLifetimeAct^[unToolNestCount] >= (parunToolLifetimeSet^[unToolNestCount] * 100)				(* Tool lifetime was exceeded *)
	THEN
		IF paretToolStatus^[unToolNestCount] = ET_ToolStatus_eOk										(* Satus is OK *)
		THEN
			paretToolStatus^[unToolNestCount] := ET_ToolStatus_eLifettimeExceeded;						(* Tool lifetime exceeded *)
			bToolLifetimeReached := TRUE; 														(* Tool lifetime reached *)
		END_IF
	END_IF;
END_IF;

IF paretToolStatus^[unToolNestCount] = ET_ToolStatus_eLifettimeExceeded								(* Tool lifetime exceeded *)
     AND (
		parunToolLifetimeSet^[unToolNestCount] = 0													(* If 0 then tool lifetime monitoring is not active *)
      		OR ((parunToolLifetimeSet^[unToolNestCount] * 100) > parunToolLifetimeAct^[unToolNestCount])  			(* Tool lifetime not exceeded *)
    	       )
THEN
	paretToolStatus^[unToolNestCount] := ET_ToolStatus_eOk;											(* Tool Ok *)
END_IF


(* Measurement tool lifetime *)
IF bToolLifetimeOn
THEN
	(* Save tool lifetime with tool change *)
	IF unToolNestAct <> unLifetimeOnNewTool				(* New tool in came *)
	    OR (
			bToolLifetimeReached							(* Tool lifetime reached *)
			AND parunToolLifetimeAct^[unToolNestAct] = 0
		  )
	THEN
		unLifetimeOnNewTool := unToolNestAct ;
		rToolLifetime := parunToolLifetimeAct^[unToolNestAct];
		bToolLifetimeReached := FALSE; 					(* Tool lifetime reached *)
	END_IF

	(*rToolLifetime:=  rToolLifetime +(rToolRotationalSpeedAct * UDINT_TO_REAL(SystemTaskInfoArr[1].cycleTime) / 100000000);*)

	rToolLifetime :=  rToolLifetime +(rToolRotationalSpeedAct * lrTaskCycle);

	IF unToolNestAct <> 0
	THEN
		parunToolLifetimeAct^[unToolNestAct] := REAL_TO_UINT(rToolLifetime);
	END_IF

END_IF


(* Reset selected tool nests *)
rtResetSelectedToolNest(
	CLK := bResetSelectedToolNest
);

IF rtResetSelectedToolNest.Q
THEN
	parunToolLifetimeAct^[unSelectedToolNest] := 0;			(* Tool lifetime clear *)

	IF parunToolNo^[unSelectedToolNest] <>  0
	THEN
		paretToolStatus^[unSelectedToolNest] := ET_ToolStatus_eOk;		(* Set tool status *)
	END_IF
END_IF;


(* Reset all tool nests *)
rtResetAllToolNests(
	CLK := bResetAllToolNests
);

IF rtResetAllToolNests.Q
THEN
	FOR unIdxToolNestCount := 1 TO unToolNestUsingMax
	DO
		IF unIdxToolNestCount <> unToolNestAct
		THEN
			parunToolLifetimeAct^[unIdxToolNestCount] := 0;			(* Tool lifetime clear *)
	
			IF parunToolNo^[unIdxToolNestCount] <>  0
			THEN
				paretToolStatus^[unIdxToolNestCount] := ET_ToolStatus_eOk;			(* Set tool status 1 = Ok*)
			END_IF
		END_IF
	END_FOR
END_IF;

(* Reset *)
IF bReset
     AND bError
THEN
	bError := FALSE;
END_IF

(* Search tool nest *)
rtExeToolNest(CLK := bExeToolNest);

IF rtExeToolNest.Q
THEN
	etToolStorage := ET_ToolStorage_eWaitExecute;                      						(* Next step *)
END_IF;

CASE etToolStorage OF
        
	ET_ToolStorage_eWaitExecute:
		bBusy := FALSE;                                     	(* Program not busy *)
		bError := FALSE;                         		(* Program not error *)
		udnErrorNo := 0;                         		(* Error number *)

		IF rtExeToolNest.Q
		THEN
			bDone := FALSE;                          	(* Program not done *)
			bBusy := TRUE;                                  (* Program busy *)

			tonWatchdog(IN := FALSE);

			unToolNestSearchCount := 0;		(* Reset tool search counter *)

			IF unToolNo = 0												(* Get old tool nest *)
			THEN
				etToolStorage := ET_ToolStorage_eGetOldToolNest;			(* Next step *)

			ELSIF unToolNo = 1000										(* Check tool place *)
			THEN
				etToolStorage := ET_ToolStorage_eChkToolPlace;			(* Next step *)

			ELSIF unToolNo = 1001										(* Check tool put up *)
			THEN
				etToolStorage := ET_ToolStorage_eChkToolPickUp;			(* Next step *)

			ELSE														(* Get new tool nest  *)
				etToolStorage := ET_ToolStorage_eGetNewToolNest;			(* Next step *)
			END_IF

		END_IF

	ET_ToolStorage_eGetNewToolNest:

			unToolNestSearchCount := unToolNestSearchCount + 1;

			IF unToolNestSearchCount <= unToolNestUsingMax
			THEN
				IF parunToolNo^[unToolNestSearchCount] = unToolNo													(* Correct tool nest found *)
				      AND (parbToolNestPresent^[unToolNestSearchCount]													(* Current nest busy *)
					        OR parunToolNo^[unToolNestSearchCount] = parunToolNo^[unToolNestUsing])						(* Identical tool number *)
				      AND paretToolStatus^[unToolNestSearchCount] = ET_ToolStatus_eOk										(* Tool status is Ok *)
				      AND ((parunToolLifetimeSet^[unToolNestSearchCount] * 100) >= parunToolLifetimeAct^[unToolNestSearchCount])		(* Tool lifetime not exceeded *)
				THEN
					IF  parunToolNo^[unToolNestSearchCount] <> parunToolNo^[unToolNestUsing]									(* Different tool number *)
				 	THEN
						IF NOT parbToolNestPresent^[unToolNestUsing]														(* Previous nest free *)
						THEN
							unToolNestPrv := unToolNestUsing;																(* Previous tool nest *)
							unToolNestAct := unToolNestSearchCount;														(* New tool nest *)

							etToolStorage := ET_ToolStorage_eDone;			(* Next step *)
						ELSE
							unToolNestPrv := 0;
							unToolNestAct := unToolNestSearchCount;

							etToolStorage := ET_ToolStorage_eError;			(* Next step *)
						END_IF
					ELSE																								(* Identical tool number *)
						IF unToolNestSearchCount = unToolNestUsing														(* Different nest number *)
						THEN																								(* Identical nest number *)
							IF paretToolStatus^[unToolNestUsing] <> ET_ToolStatus_eOk														(* Tool status is not Ok *)
							     OR ((parunToolLifetimeSet^[unToolNestUsing] * 100) < parunToolLifetimeAct^[unToolNestUsing])		(* Tool lifetime exceeded *)
							THEN
								IF NOT parbToolNestPresent^[unToolNestUsing]														(* Previous nest free *)
								THEN
									unToolNestPrv := unToolNestUsing;																(* Previous tool nest *)
									unToolNestAct := 0;														(* New tool nest *)
								
									etToolStorage := ET_ToolStorage_eDone;			(* Next step *)
								ELSE
									unToolNestPrv := unToolNestUsing;
									unToolNestAct := 0;
	
									etToolStorage := ET_ToolStorage_eError;			(* Next step *)
								END_IF
							ELSE
								(*unToolNestPrv := 0;
								unToolNestAct := unToolNestSearchCount;
	
								etToolStorage := ET_ToolStorage_eDone;			(* Next step *)*);
							END_IF
						ELSE
							IF NOT parbToolNestPresent^[unToolNestUsing]														(* Previous nest free *)
							THEN
								unToolNestPrv := unToolNestUsing;																(* Previous tool nest *)
								unToolNestAct := unToolNestSearchCount;														(* New tool nest *)

								etToolStorage := ET_ToolStorage_eDone;			(* Next step *)
							ELSE
								unToolNestPrv := 0;
								unToolNestAct := unToolNestSearchCount;
	
								etToolStorage := ET_ToolStorage_eError;			(* Next step *)
							END_IF
						END_IF
					END_IF
				END_IF
			ELSE
				IF NOT parbToolNestPresent^[unToolNestUsing]														(* Previous nest free *)
				THEN
					IF unToolNestUsing > 0
					THEN
						unToolNestPrv := unToolNestUsing;
						unToolNestAct := 0;
					END_IF

					etToolStorage := ET_ToolStorage_eError;			(* Next step *)

				ELSE
					etToolStorage := ET_ToolStorage_eError;			(* Next step *)

				END_IF
			END_IF

	ET_ToolStorage_eGetOldToolNest:
		IF NOT parbToolNestPresent^[unToolNestUsing]														(* Previous nest free *)
		THEN
			IF unToolNestUsing > 0
			THEN
				unToolNestPrv := unToolNestUsing;
				unToolNestAct := 0;
			END_IF

			etToolStorage := ET_ToolStorage_eDone;		(* Next step *)

		ELSE
			etToolStorage := ET_ToolStorage_eError;			(* Next step *)

		END_IF

	ET_ToolStorage_eChkToolPlace:
		tonWatchdog(
			IN := TRUE,
			PT:= tWatchdog
		);

		IF parbToolNestPresent^[unToolNestPrv]
		THEN
			tonWatchdog(IN := FALSE);

			unToolNestPrv := 0;
			unToolNestUsing := 0;

			etToolStorage := ET_ToolStorage_eDone;		(* Next step *)

		ELSIF tonWatchdog.Q
		THEN
			tonWatchdog(IN := FALSE);

			etToolStorage := ET_ToolStorage_eError;			(* Next step *)

		END_IF

	ET_ToolStorage_eChkToolPickUp:
		tonWatchdog(
			IN := TRUE,
			PT:= tWatchdog
		);

		IF NOT parbToolNestPresent^[unToolNestAct]
		THEN
			tonWatchdog(IN := FALSE);

			unToolNestUsing := unToolNestAct;

			etToolStorage := ET_ToolStorage_eDone;		(* Next step *)

		ELSIF tonWatchdog.Q
		THEN
			tonWatchdog(IN := FALSE);

			etToolStorage := ET_ToolStorage_eError;			(* Next step *)

		END_IF

	ET_ToolStorage_eDone:
		bDone := TRUE;				(* Program done *)
		bBusy := FALSE;                                (* Program not busy *)

		etToolStorage := ET_ToolStorage_eNoExecute;            (* Next step *)

	ET_ToolStorage_eError:
	         bDone := FALSE;				(* Program not done *)
	         bError := TRUE;				(* Program error  *)
	         bBusy := FALSE;				(* Program not busy *)

		etToolStorage := ET_ToolStorage_eNoExecute;            (* Next step *)

	ET_ToolStorage_eNoExecute:
		IF NOT bExeToolNest
		THEN
			bDone := FALSE;			(* Program not done *)
			bBusy := FALSE;                       (* Program not busy *)
			bError := FALSE;                       (* Program not error *)
			udnErrorNo := 0;                        (* Error number *)

			etToolStorage := ET_ToolStorage_eWaitExecute;              (* Next step *)

		END_IF;
END_CASE;

END_FUNCTION_BLOCK

// ---- POUs/Tc2 Objects/Automation/Spindle/FB_VFD_SpindlePreheat.TcPOU
FUNCTION_BLOCK FB_VFD_SpindlePreheat
(*

The function block used to start spindle preheat procedure.

Constructor: 		Patryk Panylo
Company:		E. Riexinger GmbH
Date:			26.06.2015
Version:			1.00

Date:			Revision:		Who:				Comment
dd.mm.yyyy		x.xx			Initials			comment

*)
VAR_INPUT
	(* Input variables / Eingang Variablen *)
	bEnable						:BOOL;						(* Enable FB signal *)
	bNoEmergencyStop			:BOOL;						(* NotAus signal *)
	bExecute					:BOOL;						(* Spindle start *)
	bInterrupt						:BOOL;						(* Interrupt *)
	bPlusRelease				:BOOL;						(* Plus move release *)
	bMinusRelease				:BOOL;						(* Minus move release *)
	bReset						:BOOL;						(* Reset procedure*)
	bCtrlEnabled					:BOOL;						(* Controller enabled *)
	bSetNewSpdlPreheat			:BOOL;						(* Set new spindle preheat *)
	bSetDailyPreheat				:BOOL;						(* Set daily preheat *)
	tSetPeriod					:TIME;						(* Set period time *)
	lrToolLimitMax				:LREAL;						(* Max rpm [U/min]  *)
	lrSpeedLimitMax				:LREAL;						(* Max rpm [U/min]  *)
	bRpmIsZero					:BOOL;						(* Spindle standstill *)
	bRpmReached				:BOOL;						(* Spindle speed reached *)
END_VAR
VAR_OUTPUT
	(* Output variables / Ausgang Variablen *)
	bValid						:BOOL;						(* Preheat valid *)
	unSpindleDurationPercent		:UINT;						(* Actual spindle duration in percent*)
	bControlerOn					:BOOL;						(* Controler on *)
	bDone						:BOOL;						(* Program done *)
	bBusy						:BOOL;						(* Program busy *)
	bError						:BOOL;						(* Program error *)
	udnErrorNo					:UDINT;						(* Error number *)
	sErrorMsg					:STRING;
END_VAR
VAR_IN_OUT
	(* Input Output variables / Ausgang Variablen *)
	Axis							:ST_VFD_AXIS_REF;					(* The AXIS_REF data type  is an interface between the PLC and the NC and contains axis information *)
	arstPhasesNewSpdl			:ARRAY [1..ungGr05MaxPhasesNewSpdl] OF ST_SpindlePreheat; 				(* Starting new spindel phases *)
	arstPhasesDailyPreheat		:ARRAY [1..ungGr05MaxPhasesDailyPreheat] OF ST_SpindlePreheat; 			(* Starting daily preheat phases *)
END_VAR
VAR
	(* Enummerations *)
	etSpindlePreheat				:ET_SpindlePreheat;				(* Spindle  mode enum variable *)

	(* Variables *)
	otstTime						:OTSTRUCT;						(* Time in OTSTRUCT *)
	unPhase						:UINT;							(* Phase counter *)
	lrSpdlTimeAsHour				:LREAL;							(* The running time of spindle procedures [h] *)
	lrStartSpdlProcTimeAsHour		:LREAL;							(* Start time of spindle procedure [h] *)
	lrSystemNewTimeAsHour 		:LREAL; 							(* System Time [h] *)
	lrPeriodAsHour				:LREAL; 							(* Period Time [h] *)
	lrWeekAsHour				:LREAL;							(* Week [h] *)
	lrDayAsHour					:LREAL;							(* Day [h] *)
	lrHour						:LREAL;							(* Hour [h] *)
	lrMinuteAsHour				:LREAL;							(* Minute Time [h] *)
	lrSecondAsHour				:LREAL;							(* Second Time [h] *)
	lrMillisecondAsHour			:LREAL;							(* Millisecond Time [h] *)

	bNewSpdl					:BOOL; 							(* New spindel phases *)
	bDailyPreheat				:BOOL; 							(* Daily preheat phases *)

	bFirstTime					:BOOL;

	(* References *)

	(* Interfaces *)

	(* Instances *)
	fbGetSystemTime				:GETSYSTEMTIME;				(* Detects System time *)
	rtReset						:R_TRIG; 						(* Positive edge for reset procedure *)
	rtExecute						:R_TRIG;							(* Positive edge for execute *)
	tonDuration					:TON;
	fbMoveVelo					:FB_VFD_MoveVelocity;
	fbStop						:FB_VFD_Stop;
	tonCtrlEnabled				:TON;
	rtSetNewSpdlPreheat			:R_TRIG;							(* Set new spindle preheat *)
	rtSetDailyPreheat				:R_TRIG;							(* Set daily preheat *)
END_VAR
VAR PERSISTENT
	lrSystemOldTimeAsHour 		:LREAL; 						(* System Time [h] *)
	bProcInterrupted				:BOOL;						(* Statring procedure interupted *)
END_VAR


IF NOT bEnable						(* Signal FB enable *)
THEN
	bValid := FALSE;;					(* Preheat valid *)
	bControlerOn := FALSE;			(* Controler off *)
	bDone := FALSE;					(* Program done *)
	bBusy := FALSE;                                  	(* Program not busy *)
	bError := FALSE;                                 	(* Program not error *)
	udnErrorNo := 0;                                 		(* Error number *)

	tonCtrlEnabled(IN := FALSE);

	bFirstTime := FALSE;

	RETURN;
END_IF;

(* Calculate system time *)
fbGetSystemTime();
lrSystemNewTimeAsHour := UINT64_TO_LREAL(IN := ULARGE_INTEGER(
	dwHighPart := fbGetSystemTime.timeHiDW,
	dwLowPart := fbGetSystemTime.timeLoDW))
	/ 10				(* Calculate into mycro seconds *)
	/ 1000			(* Calculate into millis econds *)
	/ 1000			(* Calculate into seconds *)
	/ 60				(* Calculate into minutes *)
	/ 60;				(* Calculate into hours *)

(* Calculate period time *)
otstTime := TIME_TO_OTSTRUCT(TIN := tSetPeriod);

lrWeekAsHour := otstTime.wWeek * 168.0;						(* Calculate into hours*)
lrDayAsHour := otstTime.wDay * 24.0;							(* Calculate into hours *)
lrHour := otstTime.wHour ;
lrMinuteAsHour := otstTime.wMinute  / 60.0;						(* Calculate into hours *)
lrSecondAsHour := otstTime.wSecond / 3600.0;					(* Calculate into hours *)
lrMillisecondAsHour := otstTime.wMilliseconds / 3600000.0 ;		(* Calculate into hours *)

lrPeriodAsHour :=  lrWeekAsHour							(* Calculate period *)
				+ lrDayAsHour
				+ lrHour
				+ lrMinuteAsHour
		 		+ lrSecondAsHour
				+ lrMillisecondAsHour;

(* Save last time activated of spindle *)
IF NOT Axis.bNotMoving			(* Axis moving *)
    (*AND Axis.nCurrentMotorSpeed <> 0 *)
    AND NOT bProcInterrupted
    AND NOT bBusy
THEN
	lrSystemOldTimeAsHour := lrSystemNewTimeAsHour;
END_IF

rtSetNewSpdlPreheat(CLK := bSetNewSpdlPreheat);
rtSetDailyPreheat(CLK := bSetDailyPreheat);

IF rtSetNewSpdlPreheat.Q
THEN
	lrSystemOldTimeAsHour := 0.0;
ELSIF rtSetDailyPreheat.Q
	    AND lrSystemOldTimeAsHour <> 0
THEN
	lrSystemOldTimeAsHour := 1.0;
END_IF

rtReset (CLK := bReset);											(* Positive edge for reset procedure*)
IF rtReset.Q
     AND bError
THEN
	bControlerOn := FALSE;				(* Controler off *)
	bDone := FALSE;					(* Program done *)
	bBusy := FALSE;                                  	(* Program not busy *)
	bError := FALSE;                                 	(* Program not error *)
	udnErrorNo := 0;                                 		(* Error number *)

	(* The function block MC_MoveVelocity starts a continuous movement with specified velocity and direction.  *)
	fbMoveVelo(
		bExecute := FALSE,
		Axis := Axis,
	 );

	(* The function block MC_Stop stops an axis with a defined braking ramp and blocks the axis for any motion commands.  *)
	fbStop(
		bExecute := FALSE,
		Axis := Axis,
	);

	tonDuration(IN:= FALSE);

	etSpindlePreheat := ET_SpindlePreheat_eWaitExecute;       			(* Next step *)

END_IF

(* Positive edge for execute *)
rtExecute(CLK := bExecute);
IF rtExecute.Q
THEN
	tonCtrlEnabled(IN := FALSE);

	bControlerOn := bMinusRelease
     				   AND bPlusRelease
     				   AND bNoEmergencyStop
     				   AND NOT bInterrupt;

	IF lrSystemNewTimeAsHour - lrSystemOldTimeAsHour < lrPeriodAsHour
	THEN
		bControlerOn := FALSE;
		bValid := TRUE;
	ELSE
		bValid := FALSE;
	END_IF

	RETURN;
ELSE
	tonCtrlEnabled(IN := bControlerOn
					   AND NOT bCtrlEnabled,
				   PT := t#3s);

	IF NOT bControlerOn
	     OR NOT bCtrlEnabled
	THEN
		bBusy := FALSE;                                 	(* Program not busy *)

		IF tonCtrlEnabled.Q
		THEN
			bControlerOn := FALSE;
		END_IF

		RETURN;
	ELSE
		tonCtrlEnabled(IN := FALSE);
	END_IF
END_IF;

IF NOT bCtrlEnabled
     OR NOT bNoEmergencyStop
     OR NOT bMinusRelease
     OR NOT bPlusRelease
     OR bInterrupt
THEN
	bControlerOn := FALSE;			(* Controler off *)

	(* Interrupt only when procedure has been busy  *)
	IF bBusy
	     AND NOT bProcInterrupted
	THEN
		bBusy := FALSE;                                 	(* Program not busy *)
		bProcInterrupted := TRUE;
	END_IF

	IF Axis.bNotMoving			(* Axis not moving *)
	THEN
		unSpindleDurationPercent := 0;
	END_IF

	bFirstTime := FALSE;

	RETURN;
END_IF

IF NOT bFirstTime
THEN
	bDone := FALSE;                                	(* Program done *)
	bBusy := FALSE;                                 	(* Program not busy *)
	bError := FALSE;                                 	(* Program not error *)
	udnErrorNo := 0;                                 		(* Error number *)

	(* The function block MC_MoveVelocity starts a continuous movement with specified velocity and direction.  *)
	fbMoveVelo(
		bExecute := FALSE,
		Axis := Axis,
	 );

	(* The function block MC_Stop stops an axis with a defined braking ramp and blocks the axis for any motion commands.  *)
	fbStop(
		bExecute := FALSE,
		Axis := Axis,
	);

	tonDuration(IN:= FALSE);

	etSpindlePreheat := ET_SpindlePreheat_eWaitExecute;       			(* Next step *)

	bFirstTime := TRUE;
END_IF;

IF bBusy
     (*AND Axis.nCurrentMotorSpeed <> 0*)
     AND NOT Axis.bNotMoving			(* Axis moving *)
THEN
	IF lrSystemNewTimeAsHour - lrStartSpdlProcTimeAsHour >= lrSpdlTimeAsHour
	THEN
		lrStartSpdlProcTimeAsHour := lrSystemNewTimeAsHour;
		IF unSpindleDurationPercent < 100
		THEN
			unSpindleDurationPercent := unSpindleDurationPercent + 1;
		ELSE
			unSpindleDurationPercent := 100;
		END_IF
	END_IF
ELSE
	IF Axis.bNotMoving			(* Axis not moving *)
	THEN
		unSpindleDurationPercent := 0;
	END_IF
END_IF

CASE etSpindlePreheat OF

	ET_SpindlePreheat_eWaitExecute:
		bBusy := FALSE;                                     		(* Program not busy *)
		bError := FALSE;                                    		(* Program not error *)

		bNewSpdl := FALSE; 					(* New spindel phases *)
		bDailyPreheat := FALSE; 				(* Daily preheat phases *)

		IF bControlerOn
		    AND bCtrlEnabled
		THEN
			bDone := FALSE;						(* Command done *)
			bBusy := TRUE;						(* Command busy *)
			bError := FALSE;						(* Command error  *)
			udnErrorNo := 0;						(* Error number *)
			sErrorMsg := ''; 						(* Error message *)

			tonDuration(IN:= FALSE);
			lrSpdlTimeAsHour := 0.0;

			(* New spindle starting procedure *)
			IF lrSystemOldTimeAsHour = 0
			THEN

				FOR unPhase := 1 TO ungGr05MaxPhasesNewSpdl
				DO
					(* Convert  duration time to OTSTRUCT*)
					arstPhasesNewSpdl[unPhase].otstDuration := TIME_TO_OTSTRUCT(TIN := arstPhasesNewSpdl[unPhase].tDuration);

					(* Calculate period time *)
					lrWeekAsHour := arstPhasesNewSpdl[unPhase].otstDuration.wWeek * 168.0;						(* Calculate into hours*)
					lrDayAsHour := arstPhasesNewSpdl[unPhase].otstDuration.wDay * 24.0;							(* Calculate into hours *)
					lrHour := arstPhasesNewSpdl[unPhase].otstDuration.wHour;
					lrMinuteAsHour := arstPhasesNewSpdl[unPhase].otstDuration.wMinute  / 60.0;						(* Calculate into hours *)
					lrSecondAsHour := arstPhasesNewSpdl[unPhase].otstDuration.wSecond / 3600.0;					(* Calculate into hours *)
					lrMillisecondAsHour := arstPhasesNewSpdl[unPhase].otstDuration.wMilliseconds / 3600000.0 ;			(* Calculate into hours *)

					lrSpdlTimeAsHour :=  lrSpdlTimeAsHour														(* Calculate period *)
									      + lrWeekAsHour
									      + lrDayAsHour
							 	    	      + lrHour
									      + lrMinuteAsHour
							 	    	      + lrSecondAsHour
									      + lrMillisecondAsHour;

					(* Set Limited Override *)
					arstPhasesNewSpdl[unPhase].dwOverride := LIMIT(
						0,														(* Min 0 [%]  override*)
						arstPhasesNewSpdl[unPhase].dwOverride,					(* Current [%] override*)
						100														(* Max 100 [%] override *)
					);

					(* Set Speed *)
					arstPhasesNewSpdl[unPhase].dwSpeedRpm := (LREAL_TO_DWORD(lrToolLimitMax) * arstPhasesNewSpdl[unPhase].dwOverride)/100;				(* Current RPM [U/min] *)

				END_FOR

				lrSpdlTimeAsHour := lrSpdlTimeAsHour / 100.0; 				(* Normalized to [%]*)
				lrStartSpdlProcTimeAsHour := lrSystemNewTimeAsHour;

				unPhase := 1;
				bBusy := TRUE;				(* Program Busy *)
				bNewSpdl := TRUE; 					(* New spindel phases *)
				bProcInterrupted := FALSE;

				etSpindlePreheat := ET_SpindlePreheat_eStartNewSpindle;		(* Next step *)

			(* Daily preheat starting procedure *)
			ELSIF lrSystemNewTimeAsHour - lrSystemOldTimeAsHour > lrPeriodAsHour
			THEN

				FOR unPhase := 1 TO ungGr05MaxPhasesDailyPreheat
				DO
					(* Convert  duration time to OTSTRUCT*)
					arstPhasesDailyPreheat[unPhase].otstDuration := TIME_TO_OTSTRUCT(TIN := arstPhasesDailyPreheat[unPhase].tDuration);

					(* Calculate period time *)
					lrWeekAsHour := arstPhasesDailyPreheat[unPhase].otstDuration.wWeek * 168.0;						(* Calculate into hours*)
					lrDayAsHour := arstPhasesDailyPreheat[unPhase].otstDuration.wDay * 24.0;							(* Calculate into hours *)
					lrHour := arstPhasesDailyPreheat[unPhase].otstDuration.wHour ;
					lrMinuteAsHour := arstPhasesDailyPreheat[unPhase].otstDuration.wMinute  / 60.0;						(* Calculate into hours *)
					lrSecondAsHour := arstPhasesDailyPreheat[unPhase].otstDuration.wSecond / 3600.0;					(* Calculate into hours *)
					lrMillisecondAsHour := arstPhasesDailyPreheat[unPhase].otstDuration.wMilliseconds / 3600000.0 ;			(* Calculate into hours *)

					lrSpdlTimeAsHour :=  lrSpdlTimeAsHour															(* Calculate period *)
									     + lrWeekAsHour
									     + lrDayAsHour
							 	    	     + lrHour
									     + lrMinuteAsHour
							 	   	     + lrSecondAsHour
									     + lrMillisecondAsHour;

					(* Set Limited Override *)
					arstPhasesDailyPreheat[unPhase].dwOverride := LIMIT(
						0,														(* Min 0 [%]  override*)
						arstPhasesDailyPreheat[unPhase].dwOverride,				(* Current [%] override*)
						100														(* Max 100 [%] override *)
					);

					(* Set Speed *)
					arstPhasesDailyPreheat[unPhase].dwSpeedRpm := (LREAL_TO_DWORD(lrToolLimitMax) * arstPhasesDailyPreheat[unPhase].dwOverride)/100;				(* Current RPM [U/min] *)

				END_FOR

				lrSpdlTimeAsHour := lrSpdlTimeAsHour / 100.0; 				(* Normalized to [%]*)
				lrStartSpdlProcTimeAsHour := lrSystemNewTimeAsHour;

				unPhase := 1;
				bBusy := TRUE;				(* Program Busy *)
				bDailyPreheat := TRUE; 				(* Daily preheat phases *)
				bProcInterrupted := FALSE;

				etSpindlePreheat := ET_SpindlePreheat_eStartDailyPreheat;		(* Next step *)

			END_IF;
		END_IF;

	ET_SpindlePreheat_eStartNewSpindle:
		fbMoveVelo.lrVelocity := arstPhasesNewSpdl[unPhase].dwSpeedRpm;				(* Set speed RPM [U/min] *)
		tonDuration.PT := arstPhasesNewSpdl[unPhase].tDuration;							(* Set duration time *)

		etSpindlePreheat := ET_SpindlePreheat_eStartSpindle;		(* Next step *)

	ET_SpindlePreheat_eStartDailyPreheat:
		fbMoveVelo.lrVelocity := arstPhasesDailyPreheat[unPhase].dwSpeedRpm;			(* Set speed RPM [U/min] *)
		tonDuration.PT := arstPhasesDailyPreheat[unPhase].tDuration;						(* Set duration time *)

		etSpindlePreheat := ET_SpindlePreheat_eStartSpindle;		(* Next step *)

	ET_SpindlePreheat_eStartSpindle:
		fbMoveVelo.bExecute := TRUE;

		IF fbMoveVelo.bBusy
		THEN
			etSpindlePreheat := ET_SpindlePreheat_eWfStartSpindle;         		(* Next step *)

		ELSIF fbMoveVelo.bError
		THEN
			fbMoveVelo.bExecute := FALSE;

			etSpindlePreheat := ET_SpindlePreheat_eError;         		(* Next step *)

		END_IF

	ET_SpindlePreheat_eWfStartSpindle:
		IF fbMoveVelo.bInVelocity
		     AND NOT fbMoveVelo.bError
		     AND bRpmReached
		THEN
			fbMoveVelo.bExecute := FALSE;

			etSpindlePreheat := ET_SpindlePreheat_eWfStartSpindleProc;         		(* Next step *)

		ELSIF fbMoveVelo.bError
		THEN
			fbMoveVelo.bExecute := FALSE;

			etSpindlePreheat := ET_SpindlePreheat_eError;         		(* Next step *)

		END_IF

	ET_SpindlePreheat_eWfStartSpindleProc:
		tonDuration(IN := TRUE);

		IF tonDuration.Q
		THEN
			tonDuration(IN:= FALSE);

			(* Phase incrementation *)
			unPhase := unPhase + 1;

			IF bNewSpdl
			    AND unPhase <= ungGr05MaxPhasesNewSpdl
			THEN
				fbMoveVelo.lrVelocity := arstPhasesNewSpdl[unPhase].dwSpeedRpm;				(* Set speed RPM [U/min] *)
				tonDuration.PT := arstPhasesNewSpdl[unPhase].tDuration;							(* Set duration time *)

				etSpindlePreheat := ET_SpindlePreheat_eStartSpindle;

			ELSIF bDailyPreheat
				   AND unPhase <= ungGr05MaxPhasesDailyPreheat
			THEN
				fbMoveVelo.lrVelocity := arstPhasesDailyPreheat[unPhase].dwSpeedRpm;			(* Set speed RPM [U/min] *)
				tonDuration.PT := arstPhasesDailyPreheat[unPhase].tDuration;						(* Set duration time *)

				etSpindlePreheat := ET_SpindlePreheat_eStartSpindle;

			ELSE
				etSpindlePreheat := ET_SpindlePreheat_eSpindleStop;

			END_IF
		END_IF

	ET_SpindlePreheat_eSpindleStop:
		fbStop.bExecute := TRUE;
		fbMoveVelo.lrVelocity := 0.0;

		IF fbStop.bBusy
		THEN
			etSpindlePreheat := ET_SpindlePreheat_eWfSpindleStopped;         		(* Next step *)

		ELSIF fbStop.bError
		THEN
			fbStop.bExecute := FALSE;

			etSpindlePreheat := ET_SpindlePreheat_eError;         		(* Next step *)

		END_IF

	ET_SpindlePreheat_eWfSpindleStopped:
		IF fbStop.bDone
		     AND NOT fbStop.bError
		     AND Axis.bNotMoving
		     AND Axis.nSetMotorSpeed = 0
		     AND bRpmIsZero
		THEN
			fbStop.bExecute := FALSE;

			etSpindlePreheat := ET_SpindlePreheat_eDone;         		(* Next step *)

		ELSIF fbStop.bError
		THEN
			fbStop.bExecute := FALSE;

			etSpindlePreheat := ET_SpindlePreheat_eError;         		(* Next step *)

		END_IF

	ET_SpindlePreheat_eDone:
		bValid := TRUE;						(* Preheat valid *)
		bControlerOn := FALSE;				(* Controler off *)
		bDone := TRUE;                                     		(* Program done, in position *)
		bBusy := FALSE;                                     		(* Program not busy *)

		(* Save last time activated of the starting procedure *)
		lrSystemOldTimeAsHour := lrSystemNewTimeAsHour;

		etSpindlePreheat := ET_SpindlePreheat_eNoExecute;            	(* Next step *)

	ET_SpindlePreheat_eError:
		bDone := FALSE;                                     		(* Program done, in position *)
		bControlerOn := FALSE;				(* Controler off *)
		bError := TRUE;                                     		(* Program error *)
		bBusy := FALSE;                                     		(* Program not busy *)
	
		etSpindlePreheat := ET_SpindlePreheat_eNoExecute;           	(* Next step *)

	ET_SpindlePreheat_eNoExecute:
		IF NOT bExecute
		THEN
			bNewSpdl := FALSE; 				(* New spindel phases *)
			bDailyPreheat := FALSE; 			(* Daily preheat phases *)

			bControlerOn := FALSE;				(* Controler off *)
			bDone := FALSE;                                 	(* Program done *)
			bBusy := FALSE;                                		(* Program not busy *)
			bError := FALSE;                                		(* Program not error *)
		
			etSpindlePreheat := ET_SpindlePreheat_eWaitExecute;       (* Next step *)
		
		END_IF;

END_CASE;

(* The function block MoveVelocity starts a continuous movement with specified velocity and direction.  *)
fbMoveVelo(
	lrVelocityMax := lrSpeedLimitMax,
	Axis := Axis
 );

(* The function block Stop stops an axis with a defined braking ramp and blocks the axis for any motion commands.  *)
fbStop(
	Axis := Axis,
);

END_FUNCTION_BLOCK

// ---- POUs/Tc2 Objects/Automation/Spindle/F_SpindleHSDClutchStatus.TcPOU
FUNCTION F_SpindleHSDClutchStatus : BYTE
(*

The function used to get clutch status.
.0 - Clutch is closed without tool
.1 - Clutch is closed with tool
.2 - Tool is wrong closed in clutch
.3 -  Clutch open and with tool

Constructor: 		Patryk Panylo
Company:		E. Riexinger GmbH
Date:			04.08.2015
Version:			1.00

Date:			Revision:		Who:				Comment
dd.mm.yyyy		x.xx			Initials			comment

*)
VAR_INPUT
	(* Input variables / Eingang Variablen *)
	nClutchStatus 						:INT;						(* AIx.x Status of bit clutch / Spannzange status *)
END_VAR
VAR
	(* Variables *)
	fbScaling						:FB_Scaling;
END_VAR


fbScaling(
	bEnable := TRUE,
	lrInput := INT_TO_LREAL(nClutchStatus),
	lrXLowLimit := 0,
	lrXUpperLimit := 32767,
	lrYLowLimit := 0,
	lrYUpperLimit := 10,
	usiPrecision := 2
);

F_SpindleHSDClutchStatus := 16#0;

IF fbScaling.lrOutputPV >= 5.3
     AND fbScaling.lrOutputPV <= 7.0
THEN
	F_SpindleHSDClutchStatus.0 := TRUE;			(* Clutch is closed without tool *)

ELSIF fbScaling.lrOutputPV >= 3.8
     	    AND fbScaling.lrOutputPV < 5.3
THEN
	F_SpindleHSDClutchStatus.1 := TRUE;			(* Clutch is closed with tool *)

ELSIF fbScaling.lrOutputPV >= 1.4
     	    AND fbScaling.lrOutputPV < 3.8
THEN
	F_SpindleHSDClutchStatus.2 := TRUE;			(* Tool is wrong closed in clutch *)

ELSIF fbScaling.lrOutputPV >= 1.0
     	    AND fbScaling.lrOutputPV < 1.4
THEN
	F_SpindleHSDClutchStatus.3 := TRUE;			(* Clutch without tool *)

END_IF

END_FUNCTION

// ---- POUs/Tc2 Objects/Automation/Spindle/F_SpindlePDSXLA170ClutchStatus.TcPOU
FUNCTION F_SpindlePDSXLA170ClutchStatus : ET_SpindleClutchStatus
(*

The function used to get clutch status.

Constructor: 		Patryk Panylo
Company:		E. Riexinger GmbH
Date:			18.05.2018
Version:			1.00

Date:			Revision:		Who:				Comment
dd.mm.yyyy		x.xx			Initials			comment

*)
VAR_INPUT
	(* Input variables / Eingang Variablen *)
	stClutchStatus					:ST_SpindlePDSXLA170ClutchStatus; (* Clutch status  *)
END_VAR
VAR
	(* Variables *)

END_VAR


IF stClutchStatus.bRotatingS1 AND (stClutchStatus.bToolNotClampedS2 OR NOT stClutchStatus.bToolPresentS3 OR NOT stClutchStatus.bClutchInBaseS4)			(* Clutch rotating and not closed *)
THEN
	F_SpindlePDSXLA170ClutchStatus := ET_SpindleClutchStatus_RotatingNoClosed;

ELSIF NOT stClutchStatus.bToolNotClampedS2 AND NOT stClutchStatus.bToolPresentS3 AND stClutchStatus.bClutchInBaseS4			(* Clutch is closed without tool *)
THEN
	F_SpindlePDSXLA170ClutchStatus := ET_SpindleClutchStatus_ClosedWithoutTool;

ELSIF NOT stClutchStatus.bToolNotClampedS2 AND stClutchStatus.bToolPresentS3 AND stClutchStatus.bClutchInBaseS4				(* Clutch is closed with tool *)
THEN
	F_SpindlePDSXLA170ClutchStatus := ET_SpindleClutchStatus_ClosedWithTool;

ELSIF stClutchStatus.bToolNotClampedS2 AND NOT stClutchStatus.bToolPresentS3 AND NOT stClutchStatus.bClutchInBaseS4		(* Clutch is opened *)
THEN
	F_SpindlePDSXLA170ClutchStatus := ET_SpindleClutchStatus_Opened;

ELSE
	F_SpindlePDSXLA170ClutchStatus := ET_SpindleClutchStatus_NoDefined;
END_IF

END_FUNCTION

// ---- POUs/Tc2 Objects/Automation/Spindle/F_SpindlePDSXLHClutchStatus.TcPOU
FUNCTION F_SpindlePDSXLHClutchStatus : ET_SpindleClutchStatus
(*

The function used to get clutch status.

Constructor: 		Patryk Panylo
Company:		E. Riexinger GmbH
Date:			18.05.2018
Version:			1.00

Date:			Revision:		Who:				Comment
dd.mm.yyyy		x.xx			Initials			comment

*)
VAR_INPUT
	(* Input variables / Eingang Variablen *)
	stClutchStatus						:ST_SpindlePDSXLHClutchStatus; (* Clutch status  *)
END_VAR
VAR
	(* Variables *)

END_VAR


IF NOT stClutchStatus.bSpindleStandstillS3 AND (NOT stClutchStatus.bToolClampedS1 OR stClutchStatus.bToolEjectedS2)			(* Clutch rotating and not closed *)
THEN
	F_SpindlePDSXLHClutchStatus := ET_SpindleClutchStatus_RotatingNoClosed;

ELSIF NOT stClutchStatus.bToolClampedS1 AND NOT stClutchStatus.bToolEjectedS2			(* Clutch is closed without tool *)
THEN
	F_SpindlePDSXLHClutchStatus := ET_SpindleClutchStatus_ClosedWithoutTool;

ELSIF stClutchStatus.bToolClampedS1 AND NOT stClutchStatus.bToolEjectedS2			(* Clutch is closed with tool *)
THEN
	F_SpindlePDSXLHClutchStatus := ET_SpindleClutchStatus_ClosedWithTool;

ELSIF NOT stClutchStatus.bToolClampedS1 AND stClutchStatus.bToolEjectedS2			(* Clutch is opened *)
THEN
	F_SpindlePDSXLHClutchStatus := ET_SpindleClutchStatus_Opened;

ELSE
	F_SpindlePDSXLHClutchStatus := ET_SpindleClutchStatus_NoDefined;

END_IF

END_FUNCTION

// ---- POUs/Tc2 Objects/Automation/Vacuum/FB_Vacuum.TcPOU
FUNCTION_BLOCK FB_Vacuum
(*
Base class of vacuum.

Constructor: 		Patryk Panylo
Company:		E. Riexinger GmbH
Date:			13.05.2016
Version:			1.01

Date:			Revision:		Who:				Comment
27.10.2016		.01				PPA					Monitoring of pump engine


*)
VAR_INPUT
	(* Input variables / Eingang Variablen *)
	bEnable						:BOOL;			(* Signal FB enable *)
	bAirPressure					:BOOL;			(*  Signal air pressure *)
	bEngineOk					:BOOL;			(*  Pump engine is ok *)
	bReset						:BOOL;			(*  Signal reset *)
	bAutoHand 					:BOOL;			(*  Auto := TRUE, Hand := FALSE *)
	bHandOpen					:BOOL;			(*  Hand open *)
	bHandClose					:BOOL;			(*  Hand close *)
	bAutoOpen					:BOOL;			(*  Auto open *)
	bAutoClose					:BOOL;			(*  Auto close *)
	bOpened					:BOOL;			(* Valve opened *)
	bClosed						:BOOL;			(* Valve closed *)
	bOpenRelease 				:BOOL;			(* Open release *)
	bCloseRelease				:BOOL;			(* Close release *)
	bControlStateOn				:BOOL;			(* TRUE - control with input state *)
	bControlOff					:BOOL;			(* TRUE - controle off *)
	tControlOff					:TIME;			(* Time > 0 delay to control off *)
	bValveErrOff					:BOOL;			(* TRUE -  valve off if error *)
	bErrorOff						:BOOL;			(* TRUE - error diagnose off *)
	tTimeOut						:TIME := T#5s;	(* TimeOut *)
END_VAR
VAR_OUTPUT
	(* Output variables / Ausgang Variablen *)
	bOpen						:BOOL;			(* Valve open *)
	bClose						:BOOL;			(* Valve close *)
	bEndOpened					:BOOL;			(* Open reached *)
	bEndClosed					:BOOL;			(* Close reached *)
	bNoEndPos					:BOOL;			(* End position not reached *)
	bError						:BOOL;			(* Error *)
	udnErrorNo					:UDINT;			(* Error number *)
	sErrorMsg					:STRING;		(* Error message *)

END_VAR
VAR_IN_OUT
	(* Input Output variables / Ausgang Variablen *)
	bHomeCompleted				:BOOL;			(* Home completed *)
END_VAR
VAR
	tonWatchDog					:TON;
	rtHandOpen					:R_TRIG;
	rtHandClose					:R_TRIG;
	rtAutoOpen					:R_TRIG;
	rtAutoClose					:R_TRIG;
	tonControlOff					:TON;
	bTargetOpen					:BOOL;
	bTargetClose					:BOOL;
	bFirstTime					:BOOL;

END_VAR


IF NOT bEnable
THEN
	bOpen := FALSE;                  		(* Valve open *)
	bClose := FALSE;				(* Valve close *)
	bEndOpened := FALSE;               	(* Valve opended *)
	bEndClosed := FALSE;               	(* Valve closed *)
	bError := FALSE;
	udnErrorNo := 0;                   		(* Error number *)
	sErrorMsg := '';                   		(* Error message *)

	tonWatchDog(
		IN := FALSE,
	         PT := tTimeOut
	);
	tonControlOff(
		IN := FALSE,
	         PT := tControlOff
	);

	bFirstTime := FALSE;
	RETURN;
END_IF;


IF NOT bFirstTime
THEN
	bOpen := FALSE;                    		(* Valve open *)
	bClose := FALSE;                  		(* Valve close *)
	bEndOpened := FALSE;              	(* Valve opended *)
	bEndClosed := FALSE;               	(* Valve closed *)
	bFirstTime := TRUE;
	RETURN;
END_IF;


(* Air pressure ok / Luftdruck ok *)
IF NOT bAirPressure
     OR NOT bEngineOk
THEN
	bOpen := FALSE;
	bClose := FALSE;
	bTargetOpen := FALSE;
	bTargetClose := FALSE;
	RETURN;
END_IF;


(* Check inputs  *)
rtHandOpen(CLK := bHandOpen);
rtHandClose(CLK := bHandClose);
rtAutoOpen(CLK := bAutoOpen AND bOpenRelease AND (NOT bControlOff OR tControlOff > t#0ms));
rtAutoClose(CLK := bAutoClose AND bCloseRelease AND (NOT bControlOff OR tControlOff > t#0ms));


(* Check operating mode *)
IF bAutoHand                    (* Automatic *)
THEN
	IF rtAutoOpen.Q
	    AND NOT bError
	THEN
		bTargetOpen := TRUE;
		bTargetClose := FALSE;
	END_IF;
	
	IF rtAutoClose.Q
	    AND NOT bError
	THEN
		bTargetOpen := FALSE;
		bTargetClose := TRUE;
	END_IF;
    
ELSE                        (* Manual *)
	IF rtHandOpen.Q
	   AND bOpenRelease
	   (* AND NOT #bError *)
	THEN
		bTargetOpen := TRUE;
		bTargetClose := FALSE;
	END_IF;
	
	IF rtHandClose.Q
	    AND bCloseRelease
	    (* AND NOT #bError *)
	THEN
		bTargetOpen := FALSE;
		bTargetClose := TRUE;
	END_IF;
    
END_IF;


(* Set outputs valve open *)
IF bOpenRelease
THEN
	IF bTargetOpen
	     AND NOT bOpen
	THEN
		bOpen := TRUE;
		bClose := FALSE;
		tonWatchDog(
			IN := FALSE,
			PT := tTimeOut
		);

		tonControlOff(
			IN := FALSE,
			PT := tControlOff
		);
	END_IF;
    
ELSE
	IF bTargetOpen
	    AND bOpen
	THEN
		bOpen := FALSE;
	
		IF NOT bAutoHand
		THEN
		    bTargetOpen := FALSE;
		END_IF;
	
	END_IF;
END_IF;

(* Set outputs valve close *)
IF bCloseRelease
THEN
	IF bTargetClose
	    AND NOT bClose
	THEN
		bOpen := FALSE;
		bClose := TRUE;
		tonWatchDog(
			IN := FALSE,
			PT := tTimeOut
		);

		tonControlOff(
			IN := FALSE,
			PT := tControlOff
		);
	END_IF;
    
ELSE
	IF bTargetClose
	     AND bClose
	THEN
		bClose := FALSE;

		IF NOT bAutoHand
		THEN
			bTargetClose := FALSE;
		END_IF;
	
	END_IF;
END_IF;

IF NOT bAutoHand
     AND (bOpen OR bClose)
THEN
	bHomeCompleted := FALSE;
END_IF;

(* Error reset *)
IF bReset
    AND bError
THEN
	udnErrorNo := 0;                    (* Error number *)
	sErrorMsg := '';                    (* Error message *)
	tonWatchDog(
		IN := FALSE,
	         PT := tTimeOut
	);

END_IF;

(* Timer starts when valve is not opened and work position *)
tonWatchDog(
	IN := NOT bErrorOff
		AND (
			(bClose AND NOT bClosed)
			  OR (bOpen AND NOT bOpened)
			  OR (NOT bOpened AND NOT bClosed)
			  OR (bOpened AND bClosed)),
	PT := tTimeOut
);

(* Error if valve does not reach open or work sensor *)
IF tonWatchDog.Q
    AND NOT bError
THEN
	IF bClose
	THEN
		IF NOT bClosed AND NOT bOpened
		THEN
			udnErrorNo := 1;                                (* Set error number *)
			sErrorMsg := 'Work position not reached';
		ELSIF NOT bClosed AND bOpened
		THEN
			udnErrorNo := 2;                                (* Set error number *)
			sErrorMsg := 'Not move in work position';
		ELSIF bClosed AND bOpened
		THEN
			udnErrorNo := 5;                                    (* Set error number *)
			sErrorMsg := 'Both position reached';
		END_IF;
	ELSIF bOpen
	THEN
		IF NOT bClosed AND NOT bOpened
		THEN
			udnErrorNo := 3;                                (* Set error number *)
			sErrorMsg := 'Base position not reached';
		ELSIF bClosed AND NOT bOpened
		THEN
			udnErrorNo := 4;                                (* Set error number *)
			sErrorMsg := 'Not move in base position';
		ELSIF bClosed AND bOpened
		THEN
			udnErrorNo := 5;                                    (* Set error number *)
			sErrorMsg := 'Both position reached';
		END_IF;
	ELSIF bClosed AND bOpened
	THEN
		udnErrorNo := 5;                                    (* Set error number *)
		sErrorMsg := 'Both position reached';
	END_IF;
END_IF;

bError := udnErrorNo <> 0;

(* Open reached  *)
bEndOpened := bOpened
			    AND NOT bClosed
			    AND NOT bError;

(* Close reached  *)
bEndClosed := NOT bOpened
			  AND bClosed
			  AND NOT bError;

(* End position not reached *)
IF bTargetOpen
THEN
	bNoEndPos := NOT bOpened;
    
ELSIF bTargetClose
THEN
	bNoEndPos := NOT bClosed;

ELSE
    bNoEndPos := FALSE;
END_IF;


(* Valve off if error  *)
IF bError
    AND (bOpen OR bClose)
    AND bValveErrOff
THEN
	bOpen := FALSE;
	bClose := FALSE;
END_IF;

(* Control with input state *)
IF bControlStateOn
THEN
	IF bAutoHand					(* Automatic *)
	THEN
		IF NOT bAutoOpen
		THEN
			bOpen := FALSE;
			bTargetOpen := FALSE;
		END_IF

		IF NOT bAutoClose
		THEN
			bClose := FALSE;
			bTargetClose := FALSE;
		END_IF
	
	ELSE						(* Manual *)
		IF NOT bHandOpen
		THEN
			bOpen := FALSE;
			bTargetOpen := FALSE;
		END_IF

		IF NOT bHandClose
		THEN
			bClose := FALSE;
			bTargetClose := FALSE;
		END_IF
	
	END_IF;
END_IF

(* Check control off *)
IF bControlOff
   AND tControlOff > t#0ms
THEN
	tonControlOff(
		IN := bOpen OR bClose
			 OR bTargetOpen OR bTargetClose,
		PT := tControlOff
	);
    
	IF tonControlOff.Q
	THEN
		bOpen := FALSE;
		bClose := FALSE;
		bTargetOpen := FALSE;
		bTargetClose := FALSE;
	END_IF;
    
ELSE
	tonControlOff(
		IN := FALSE,
		PT := tControlOff
	);
	
	IF bControlOff
	     AND (bOpen OR bClose
		       OR bTargetOpen OR bTargetClose)
	THEN
		bOpen := FALSE;
		bClose := FALSE;
		bTargetOpen := FALSE;
		bTargetClose := FALSE;
	END_IF;
END_IF;

END_FUNCTION_BLOCK

// ---- POUs/Tc2 Objects/Basics/FB_Get_Time.TcPOU
FUNCTION_BLOCK FB_Get_Time
VAR_INPUT
END_VAR
VAR_OUTPUT
	sDateAndTime: STRING;
END_VAR
VAR
	bBusy: BOOL;
	bError: BOOL;
	udiErrorID: UDINT;
	fbGetTime: NT_GetTime;
	stTime: TIMESTRUCT;
	nStep: UDINT;
	bBlinker: BOOL;
	fbBlinker: FB_Blinker;
	stBlinker:ST_Blinker;
END_VAR

(*This Function Block gets the Windows Systemtime*)

CASE nStep OF
	0:	IF NOT bError AND NOT bBusy THEN
			nStep:= 10;
		ELSE
			nStep:= 30;
		END_IF

	10:	IF stBlinker.Q0 THEN
			fbGetTime.START:= TRUE;
		ELSE
			fbGetTime.START:= FALSE;
			nStep:= 0;
		END_IF

	30:	IF NOT bError AND NOT bBusy THEN
			nStep:= 10;
		END_IF
END_CASE

fbBlinker(tPeriod := t#500ms, stBlinker => stBlinker);

fbGetTime(
			NETID:= '' ,
			START:=   ,
			TMOUT:= DEFAULT_ADS_TIMEOUT ,
			BUSY=> bBusy ,
			ERR=> bError ,
			ERRID=> udiErrorID ,
			TIMESTR=> stTime );

sDateAndTime:= SYSTEMTIME_TO_STRING(stTime);

END_FUNCTION_BLOCK

// ---- POUs/Tc2 Objects/Basics/F_AdsError_Text.TcPOU
FUNCTION F_AdsError_Text : STRING
VAR_INPUT
	nCode: UDINT;
END_VAR
VAR
	sText: STRING(255);
END_VAR

CASE nCode OF
	16#000 : sText := '0: No error  ';
	16#001 : sText := '1: Internal error  ';
	16#002 : sText := '2: No Rtime  ';
	16#003 : sText := '3: Allocation locked memory error  ';
	16#004 : sText := '4: Insert mailbox error  ';
	16#005 : sText := '5: Wrong receive HMSG  ';
	16#006 : sText := '6: target port not found  ';
	16#007 : sText := '7: target machine not found  ';
	16#008 : sText := '8: Unknown command ID  ';
	16#009 : sText := '9: Bad task ID  ';
	16#00A : sText := '10: No IO  ';
	16#00B : sText := '11: Unknown AMS command  ';
	16#00C : sText := '12: Win 32 error  ';
	16#00D : sText := '13: Port not connected  ';
	16#00E : sText := '14: Invalid AMS length  ';
	16#00F : sText := '15: Invalid AMS Net ID  ';
	16#010 : sText := '16: Low Installation level  ';
	16#011 : sText := '17: No debug available  ';
	16#012 : sText := '18: Port disabled  ';
	16#013 : sText := '19: Port already connected  ';
	16#014 : sText := '20: AMS Sync Win32 error  ';
	16#015 : sText := '21: AMS Sync Timeout  ';
	16#016 : sText := '22: AMS Sync AMS error  ';
	16#017 : sText := '23: AMS Sync no index map  '; 
	16#018 : sText := '24: Invalid AMS port  ';
	16#019 : sText := '25: No memory  ';
	16#01A : sText := '26: TCP send error  ';
	16#01B : sText := '27: Host unreachable  ';
	16#1000 : sText := '4096: Intern: RTERR_INTERNAL : $R$N Internal fatal error in the TwinCAT real-time system.  ';
	16#1001 : sText := '4097: Intern: RTERR_BADTIMERPERIODS: $R$N Timer value not vaild.  ';
	16#1002 : sText := '4098: Intern: RTERR_INVALIDTASKPTR: $R$N Task pointer has the invalid value ZERO. ';
	16#1003 : sText := '4099: Intern: RTERR_INVALIDSTACKPTR: $R$N Task stack pointer has the invalid value ZERO. ';
	16#1004 : sText := '4100: Intern: RTERR_PRIOEXISTS: $R$N The demand task priority is already assigned.  ';
	16#1005 : sText := '4101: Intern: RTERR_NOMORETCB: $R$N No more free TCB (Task Control Block) available. Maximum number of TCBs is 64.  ';
	16#1006 : sText := '4102: Intern: RTERR_NOMORESEMAS: $R$N No more free semaphores available. Maximum number of semaphores is 64.  ';
	16#1007 : sText := '4103: Intern: RTERR_NOMOREQUEUES: $R$N No more free queue available. Maximum number of queue is 64.  ';
	16#1008 : sText := '4104: Intern: TwinCAT reserved.:  ';
	16#1009 : sText := '4105: Intern: TwinCAT reserved.:  '; 
	16#100a : sText := '4106: Intern: TwinCAT reserved.:  '; 
	16#100b : sText := '4107: Intern: TwinCAT reserved.:  '; 
	16#100C : sText := '4108: Intern: TwinCAT reserved.:  ';
	16#100D : sText := '4109: Intern: RTERR_EXTIRQALREADYDEF: $R$N An external synchronisation interrupt is already applied. ';
	16#100E : sText := '4110: Intern: RTERR_EXTIRQNOTDEF: $R$N No external synchronsiation interrupt applied. ';
	16#100F : sText := '4111: Intern: RTERR_EXTIRQINSTALLFAILED: $R$N The apply of the external synchronisation interrupt failed. ';
	16#1010 : sText := '4112: Intern: RTERR_IRQLNOTLESSOREQUAL: $R$N Call of a service function in the wrong context.  ';
	16#2000 : sText := ': ERR_IOERRS  ';
	16#274C : sText := '10060: A socket operation was attempted to an unreachable host  ';
	16#274D : sText := '10061: A connection attempt failed because the connected party did not properly respond after a period of time, $R$N or established connection failed because connected host has failed to respond.  ';
	16#2751 : sText := '10065: No connection could be made because the target machine actively refused it  ';
	16#2900 : sText := ': ERR_DPSLAVE (ERR_IOERRS+0x900)  ';
	16#2A00 : sText := ': ERR_CP5412A2 (ERR_IOERRS+0xA00)  '; 
	16#2B00 : sText := ': ERR_ASP (ERR_IOERRS+0xB00)  '; 
	16#2C00 : sText := ': ERR_CANSLAVE (ERR_IOERRS+0xC00)  '; 
	16#2D00 : sText := ': ERR_CIF30 (ERR_IOERRS+0xD00)  '; 
	16#2E00 : sText := ': ERR_IBSSLAVE (ERR_IOERRS+0xE00)  ';
	16#3000 : sText := ': ERR_SPSERRS  '; 
	16#4000 : sText := ': ERR_NCERRS  ';
	16#500 : sText := '1280: Intern: ROUTERERR_NOLOCKEDMEMORY: $R$N No locked memory can be allocated.  ';
	16#501 : sText := '1281: Intern: ROUTERERR_RESIZEMEMORY: $R$N The size of the  router memory could not be changed. ';
	16#502 : sText := '1282: Intern: ROUTERERR_MAILBOXFULL: $R$N The Mailbox of the AmsPort has reached the maximum number of possible entries. The current sent message was abolished.  ';
	16#503 : sText := '1283: Intern: ROUTERERR_DEBUGBOXFULL: $R$N The Mailbox of the Ams debugger port has reached the maximum number of possible entries. $R$N The sent message wil not be displayed in the debug monitor.  ';
	16#504 : sText := '1284: Intern: ROUTERERR_UNKNOWNPORTTYPE :  ';
	16#505 : sText := '1285: Intern: ROUTERERR_NOTINITIALIZED: $R$N Router is not (yet) initialised.  ';
	16#506 : sText := '1286: Intern: ROUTERERR_PORTALREADYINUSE : $R$N The desired port number is already assigned. ';
	16#507 : sText := '1287: Intern: ROUTERERR_NOTREGISTERED : $R$N Ams Port not registered  ';
	16#508 : sText := '1288: Intern: ROUTERERR_NOMOREQUEUES: $R$N The maximum number of Ams Ports reached.  ';
	16#509 : sText := '1289: Intern: ROUTERERR_INVALIDPORT :  '; 
	16#50A : sText := '1290: Intern: ROUTERERR_NOTACTIVATED : $R$N TwinCAT Router not (yet) active.  ';
	16#6000 : sText := ': ERR_PLCERRS  ';
	16#0700 : sText := '1792: error class <device error>  ';
	16#7000 : sText := ': ERR_STRKERRS  '; 
	16#0701 : sText := '1793: Service is not supported by server  ';
	16#0702 : sText := '1794: invalid index group  ';
	16#0703 : sText := '1795: invalid index offset  ';
	16#0704 : sText := '1796: reading/writing not permitted  ';
	16#0705 : sText := '1797 : parameter size not correct  ';
	16#0706 : sText := '1798: invalid parameter value(s)  ';
	16#0707 : sText := '1799: device is not in a ready state  ';
	16#708 : sText := '1800: device is busy  '; 
	16#709 : sText := '1801: invalid context (must be in Windows)  ';
	16#70A : sText := '1802: out of memory  '; 
	16#70B : sText := '1803: invalid parameter value(s)  '; 
	16#70C : sText := '1804: not found (files, ...)  ';
	16#70D : sText := '1805: syntax error in command or file  '; 
	16#70E : sText := '1806: objects do not match  '; 
	16#70F : sText := '1807: object already exists  '; 
	16#710 : sText := '1808: symbol not found  '; 
	16#711 : sText := '1809: symbol version invalid  '; 
	16#712 : sText := '1810: server is in invalid state  '; 
	16#713 : sText := '1811: AdsTransMode not supported  '; 
	16#714 : sText := '1812: Notification handle is invalid  '; 
	16#715 : sText := '1813: Notification client not registered  '; 
	16#716 : sText := '1814: no more notification handles  '; 
	16#717 : sText := '1815: size for watch too big  ';
	16#718 : sText := '1816: device not initialized  ';
	16#719 : sText := '1817: device has a timeout  '; 
	16#71A : sText := '1818: query interface failed  '; 
	16#71B : sText := '1819: wrong interface required  '; 
	16#71C : sText := '1820: class ID is invalid  '; 
	16#71D : sText := '1821: object ID is invalid  '; 
	16#71E : sText := '1822: request is pending  '; 
	16#71F : sText := '1823: request is aborted  '; 
	16#720 : sText := '1824: signal warning  '; 
	16#721 : sText := '1825: invalid array index  ';
	16#722 : sText := '1826: symbol not active -> release handle and try again  ';
	16#723 : sText := '1827: access denied  ';
	16#740 : sText := '1856: Error class <client error>  ';
	16#741 : sText := '1857: invalid parameter at service  ';
	16#742 : sText := '1858: polling list is empty  '; 
	16#743 : sText := '1859: var connection already in use  ';
	16#744 : sText := '1860: invoke ID in use  ';
	16#745 : sText := '1861: timeout elapsed  ';
	16#746 : sText := '1862: error in win32 subsystem  '; 
	16#748 : sText := '1864: ads port not opened  '; 
	16#750 : sText := '1872: internal error in ads sync  ';
	16#751 : sText := '1873: hash table overflow  ';
	16#752 : sText := '1874: key not found in hash  ';
	16#753 : sText := '1875: no more symbols in cache  '; 
	16#754 : sText := '1876: invalid response received   ';
	16#755 : sText := '1877: Sync port locked: ADS-Client tries to send a ADS msg but another thread is still waiting for an ADS-response. $R$N This error occurs only if no ADS-router is installed (please install royalty free TwinCAT-CP) $R$N or the router does not know the remote ADS device (define the remote ADS partner )  ';
	16#7800 : sText := ': ERR_PRJSPECIFIC  ';
	ELSE
		sText := 'No Text for this ErrorCode available';
END_CASE;

F_AdsError_Text := sText;

END_FUNCTION

// ---- POUs/Tc2 Objects/Conversions/BitOriented/F_ConvArrBitsToWord.TcPOU
FUNCTION F_ConvArrBitsToWord : WORD
VAR_INPUT
	arrBits: ARRAY [0..15] OF BOOL;
END_VAR
VAR
END_VAR

F_ConvArrBitsToWord := 0;

END_FUNCTION

// ---- POUs/Tc2 Objects/Diagnostic/Terminal/FB_ToggleBit.TcPOU
FUNCTION_BLOCK FB_ToggleBit
VAR_INPUT
(*+++++ TxPDO Toggle +++++*)
	bToggle: BOOL;
END_VAR
VAR_OUTPUT
END_VAR
VAR
(*+++++ Toggle Bit Bridge +++++*)
	rtToggle: R_TRIG;
	ftToggle: F_TRIG;
	rCounter: REAL;
	rLastCounter: REAL;
(*+++++ Evaluation of Toggle Bits +++++*)
	tonTimer: TON;
	rToggleBitCounter: REAL;
	rUpdateTime: REAL;
END_VAR

(*This function block evaluates the Toggle Bit of the device.
Within a period of 10 seconds, is is checked how often the Toggle Bit changes it's value. *)

rtToggle(CLK:= bToggle);
ftToggle(CLK:= bToggle);

tonTimer.IN:= TRUE;
tonTimer.PT:= t#10000ms;

IF NOT tonTimer.Q THEN
	IF rtToggle.Q THEN
		rCounter:= rCounter+1;
	END_IF
	IF ftToggle.Q THEN
		rCounter:= rCounter+1;
	END_IF

	rToggleBitCounter:= rCounter;
ELSE
	rLastCounter:= rCounter;
	rUpdateTime:= 1/ (rLastCounter/10); 		(*Update Time is calculated*)
	rCounter:= 0;
	tonTimer.IN:= FALSE;
END_IF

tonTimer();

END_FUNCTION_BLOCK

// ---- POUs/Tc2 Objects/Engineering/Buffer/FB_FiFo.TcPOU
FUNCTION_BLOCK FB_FiFo
(*
FiFo buffer of strings.

Constructor: 		Patryk Panylo
Company:		E. Riexinger GmbH
Date:			14.05.2013
Version:			1.00

Date:			Revision:		Who:				Comment
dd.mm.yyyy		x.xx			Initials			comment

*)
VAR_INPUT
	bAdd				:BOOL;
	bClear				:BOOL;
	sItem				:STRING;
END_VAR
VAR_OUTPUT

END_VAR
VAR_IN_OUT
	arsBuffer				:ARRAY[0..unSize] OF STRING;			(* Circular buffer *)
END_VAR
VAR
	bNoBufferEmpty		:BOOL;									(* Buffer empty *)
	nIdx					:INT;

	rtAdd				:R_TRIG;
	rtClear				:R_TRIG;
END_VAR
VAR CONSTANT
	unSize				:UINT := 100;								(* Buffer size *)
END_VAR

(* Add date to buffor *)
rtAdd(CLK := bAdd);

IF rtAdd.Q
THEN
	FOR nIdx := unSize - 1 TO 0 BY -1
	DO
		arsBuffer[nIdx + 1] := arsBuffer[nIdx];
	END_FOR

	arsBuffer[0] := sItem;

	RETURN;
END_IF

(* Clear buffor *)
rtClear(CLK := bClear);

IF rtClear.Q
THEN
	MEMSET(ADR(arsBuffer), 0, SIZEOF(arsBuffer));
	nIdx := 0;
END_IF

END_FUNCTION_BLOCK

// ---- POUs/Tc2 Objects/Engineering/External set value generator/FB_ExtSetPoint.TcPOU
FUNCTION_BLOCK FB_ExtSetPoint
(*

The function block used to move axis with an external set value.

Constructor: 		Patryk Panylo
Company:		E. Riexinger GmbH
Date:			01.04.2015
Version:			1.00

Date:			Revision:		Who:				Comment
dd.mm.yyyy		x.xx			Initials			comment

*)
VAR_INPUT
	(* Input variables / Eingang Variablen *)
	bEnable					:BOOL;						(* Function block enable *)
	bStart					:BOOL;						(* Execute start an external set value generator with rising edge *)
	bStop					:BOOL;						(* Execute stop an external set value generator with rising edge *)
	lrPosition					:LREAL;						(* Set position from an external set value generator *)
	lrPositionOffset			:LREAL;						(* Set offset of position *)
	ePositionType 			:E_PositionType ;				(* Position type - POSITIONTYPE_ABSOLUTE or POSITIONTYPE_RELATIVE *)
	lrVelocity					:LREAL;						(* Set velocity from an external set point generator  > 0 *)
	lrAcceleration				:LREAL;						(* Set acceleration from an external set point generator > 0 *)
END_VAR
VAR_OUTPUT
	(* Output variables / Ausgang Variablen *)
	bEnabled  				:BOOL;						(* Enabled shows the current state of the external set point generator *)
	bDone					:BOOL;						(* Command done *)
	bBusy					:BOOL;						(* Command busy *)
	bError					:BOOL;						(* Command error  *)
	udnErrorNo				:UDINT;						(* Error number *)
	sErrorMsg				:STRING; 					(* Error message *)
END_VAR
VAR_IN_OUT
	Axis						:AXIS_REF;					(* The AXIS_REF data type  is an interface between the PLC and the NC and contains axis information *)
END_VAR
VAR
	(* Instances / Instanzen *)
	fbMC_ExtSetPointGenEnable			:MC_ExtSetPointGenEnable;						(* Switch on external set value generator with the function. *)
	fbMC_ExtSetPointGenDisable			:MC_ExtSetPointGenDisable;						(* Switch off external set value generator with the function. *)

	(* Enumerator  *)
	etMoveExtState						: ET_MoveExtState;								(* Current state *)

	(* General flags / Allgemeine Variablen *)
	eLastPositionType 					:E_PositionType;
	lrExtPosition							:LREAL;
	lrExtVelocity							:LREAL;
	lrExtAcceleration						:LREAL;
	dnExtDirection						:DINT;
	bImediateStop						:BOOL;
	bFirstTime							:BOOL;

END_VAR
VAR CONSTANT
	lrEPSILON				 :LREAL := 1E-6;
END_VAR

IF NOT bEnable
THEN
	bDone := FALSE;					(* Command done *)
	bBusy := FALSE;					(* Command busy *)
	bError := FALSE;					(* Command error  *)
	udnErrorNo := 0;					(* Error number *)
	sErrorMsg := ''; 					(* Error message *)

	bEnabled := FALSE;
	IF bStart
	THEN
		bEnabled := TRUE;
	END_IF;

	bFirstTime := FALSE;
	RETURN;
END_IF

IF NOT bFirstTime
THEN
	bEnabled := FALSE;

	fbMC_ExtSetPointGenEnable(Execute := FALSE, Axis:=Axis);						(* Reset FB and get Enabled status *)
	fbMC_ExtSetPointGenDisable(Execute := FALSE, Axis:=Axis); 						(* Reset FB and get Enabled status *)

	etMoveExtState := ET_MoveExtState_eWaitExecute;

	bFirstTime := TRUE;
END_IF

bImediateStop := AxisInErrorState(Axis.NcToPlc.AxisState);
IF bImediateStop
THEN
	(* Stop generator if axis is in error state *)
	lrExtVelocity := 0.0;
	lrExtAcceleration := 0.0;
	bError := TRUE;													(* Command error  *)
	udnErrorNo :=  Axis.NcToPlc.ErrorCode;								(* Error number *)
	sErrorMsg := ''; 													(* Error message *)

	etMoveExtState := ET_MoveExtState_eError;

ELSE
	(* Produce the dynamic data for the external setpoint generator interface *)
	lrExtVelocity := lrVelocity;
	lrExtAcceleration := lrAcceleration;
END_IF

lrExtPosition :=  lrPosition + lrPositionOffset;

IF lrExtVelocity = 0.0
    AND lrExtAcceleration = 0.0
THEN
	dnExtDirection := 0;				(* Stand still *)
END_IF

IF lrExtVelocity >= 0.0
THEN
	dnExtDirection := 1;				(* Positive motion *)
ELSE
	dnExtDirection := -1;				(* Negative motion *)
END_IF

CASE etMoveExtState
OF
	ET_MoveExtState_eWaitExecute:
		IF bStop
		THEN
			fbMC_ExtSetPointGenEnable(Execute := FALSE, Axis := Axis);						(* Reset FB and get Enabled status *)
			fbMC_ExtSetPointGenDisable(Execute := FALSE, Axis := Axis); 					(* Reset FB and get Enabled status *)

			bDone := FALSE;						(* Command done *)
			bBusy := TRUE;						(* Command busy *)
			bError := FALSE;						(* Command error  *)
			udnErrorNo := 0;						(* Error number *)
			sErrorMsg := ''; 						(* Error message *)

			etMoveExtState := ET_MoveExtState_eDisableExtSetPointGenerator;

		ELSIF bStart
		THEN
			fbMC_ExtSetPointGenEnable(Execute := FALSE, Axis := Axis);						(* Reset FB and get Enabled status *)
			fbMC_ExtSetPointGenDisable(Execute := FALSE, Axis := Axis); 					(* Reset FB and get Enabled status *)

			bDone := FALSE;						(* Command done *)
			bBusy := TRUE;						(* Command busy *)
			bError := FALSE;						(* Command error  *)
			udnErrorNo := 0;						(* Error number *)
			sErrorMsg := ''; 						(* Error message *)

			etMoveExtState := ET_MoveExtState_eEnableExtSetPointGenerator;

			(* Check for errors *)
			(* lrExtVelocity < lrEPSILON
			THEN
				udnErrorNo := 1;						(* Error number *)

				etMoveExtState := ET_MoveExtState_eError;
			END_IF
			IF lrExtAcceleration < lrEPSILON
			THEN
				udnErrorNo := 2;						(* Error number *)

				etMoveExtState := ET_MoveExtState_eError;
			END_IF*)
		END_IF

	ET_MoveExtState_eEnableExtSetPointGenerator:
		IF fbMC_ExtSetPointGenEnable.Enabled
		    AND NOT fbMC_ExtSetPointGenEnable.Execute
		    AND (ePositionType = eLastPositionType)
		THEN
			(* Send enable command to set the new target position but do not wait until the command has finished *)
			fbMC_ExtSetPointGenEnable.Execute := TRUE ;
			fbMC_ExtSetPointGenEnable.PositionType := ePositionType;

			etMoveExtState := ET_MoveExtState_eDone;

		ELSE
			(* Enable the set point generator *)
			fbMC_ExtSetPointGenEnable.Execute := TRUE ;
			fbMC_ExtSetPointGenEnable.PositionType := ePositionType;

			IF fbMC_ExtSetPointGenEnable.Error
			     AND NOT fbMC_ExtSetPointGenEnable.Busy
			THEN
				bError := fbMC_ExtSetPointGenEnable.Error;							(* Command error  *)
				udnErrorNo := fbMC_ExtSetPointGenEnable.ErrorID;						(* Error number *)

				etMoveExtState := ET_MoveExtState_eError;

			ELSIF fbMC_ExtSetPointGenEnable.Done
			     	    AND NOT fbMC_ExtSetPointGenEnable.Busy
			THEN
				eLastPositionType := ePositionType;

				etMoveExtState := ET_MoveExtState_eDone;
			END_IF

		END_IF

	ET_MoveExtState_eDisableExtSetPointGenerator:
		(* Call the disable external set point generator function block *)
		fbMC_ExtSetPointGenDisable(
			Execute := TRUE ,
			Axis:=Axis
		);
		
		IF fbMC_ExtSetPointGenDisable.Error
		     AND NOT fbMC_ExtSetPointGenEnable.Busy
		THEN
			fbMC_ExtSetPointGenDisable(
				Execute := FALSE ,
				Axis:=Axis
			);
		
			bError := fbMC_ExtSetPointGenDisable.Error;												(* Command error  *)
			udnErrorNo := fbMC_ExtSetPointGenDisable.ErrorID;										(* Error number *)

			etMoveExtState := ET_MoveExtState_eError;
		
		ELSIF fbMC_ExtSetPointGenDisable.Done
		     	    AND NOT fbMC_ExtSetPointGenEnable.Busy
		THEN
		
			etMoveExtState := ET_MoveExtState_eDone;
		END_IF

	ET_MoveExtState_eError:
		bBusy := FALSE;						(* Command busy *)
		bError := TRUE;						(* Command error  *)

		etMoveExtState := ET_MoveExtState_eNoExecute;

	ET_MoveExtState_eDone:
		bDone := TRUE;						(* Command done *)
		bBusy := FALSE;						(* Command busy *)

		etMoveExtState := ET_MoveExtState_eNoExecute;

	ET_MoveExtState_eNoExecute:
		IF NOT bStart
		     AND NOT bStop
		THEN
			(* Reset outputs *)
			bDone := FALSE;						(* Command done *)
			bBusy := FALSE;						(* Command busy *)
			bError := FALSE;						(* Command error  *)

			etMoveExtState := ET_MoveExtState_eWaitExecute;
		END_IF
END_CASE

(* The function is used to feed set values from an external set point generator into an axis. *)
MC_ExtSetPointGenFeed(
	Position := lrExtPosition,
	Velocity := 0.0,
	Acceleration := 0.0,
	Direction := dnExtDirection,
	Axis := Axis
);

(* Call the enable external set point generator function block *)
fbMC_ExtSetPointGenEnable(
	Position := lrPosition,
	Enabled => bEnabled,
	Axis:= Axis
 );

END_FUNCTION_BLOCK

// ---- POUs/Tc2 Objects/Engineering/Filter/FB_PT1.TcPOU
FUNCTION_BLOCK FB_PT1
(*

Function block low-pass filter (PT1)  for damping of fast alternating input-values.
K(s) = k/1+sT1  -> h(t) = k(1 - e^(-t/T1))

The Discrete-Time Integrator using Euler method: 
y(n+1) = 1/T1 * dt * (kp * xn - yn) + yn => kp * xn * dt / T1+ yn * (1 - dt / T1)

y(n+1) = kp * xn * Tcycle / T1+ yn * (1 - Tcycle / T1)
T1 = 0 =>  y(n+1) = kp * xn

Sample Time
Constructor: 		Patryk Panylo
Company:		E. Riexinger GmbH
Date:			20.03.2014
Version:			1.00

Date:			Revision:		Who:				Comment
dd.mm.yyyy		x.xx			Initials			comment

